	// Для таймера шага
	tonStepTimeout   : TON; // Таймер превышения времени шага
	xStepTimeout     : BOOL; // Время шага превышено
	xStepChanged     : BOOL; // Шаг изменился в текущем цикле
	xStepTimerEnable : BOOL; // Разрешение таймера шага
	xStepInitialized : BOOL; // Предыдущий шаг инициализирован
	
	// Для удержания предупреждений
    tpWarningHold : TP; // Удержание предупреждения для отображения
    xWarningPulse : BOOL; // Импульс нового предупреждения
	
	// ФБ группы осей
	fbReadStatus   : MC_GroupReadStatus; // Чтение состояния группы
	fbReadError    : MC_GroupReadError; // Чтение активной ошибки группы
	fbReadPosition : MC_GroupReadActualPosition; // Чтение текущей позиции группы
	fbGroupEnable  : MC_GroupEnable; // Включение группы
	fbGroupDisable : MC_GroupDisable; // Отключение группы
	fbGroupReset   : MC_GroupReset; // Сброс ошибок группы
	fbGroupSetOverride : MC_GroupSetOverride; // Live override активного и следующего движения группы

	
	fbMoveDirect : MC_MoveDirectAbsolute; // Прямое абсолютное перемещение
	fbMoveLinear : MC_MoveLinearAbsolute; // Линейное абсолютное перемещение
	fbFaultInjector : FB_AXIS_GROUP_FAULT_INJECTOR; // Изолированная инъекция библиотечной ошибки
	
	fbGroupHalt : MC_GroupHalt; // Плавная остановка группы
	fbGroupStop : MC_GroupStop; // Остановка группы
	
	stPosition : SMC_POS_REF; // Текущая позиция группы
	
	// Триггеры на команды
    rtEnable        : R_TRIG; // Фронт команды включения
    rtDisable       : R_TRIG; // Фронт команды отключения
	rtEnablePower   : R_TRIG; // Фронт запроса питания
    rtResetAllError : R_TRIG; // Фронт команды сброса
    rtMoveDirect    : R_TRIG; // Фронт прямого перемещения
    rtMoveLinear    : R_TRIG; // Фронт линейного перемещения
	rtStopCmd       : R_TRIG; // Фронт команды остановки
	rtHaltCmd       : R_TRIG; // Фронт плавной остановки
	
END_VAR
VAR_IN_OUT
	AxisGroup : AXIS_GROUP_REF_SM3; // Ссылка на группу осей SoftMotion
	GroupData : ST_AXIS_GROUP; // Команды, статусы и диагностика группы
END_VAR

VAR CONSTANT
	// ==================================================
    // Логические ошибки группы
    // ==================================================
	LOG_STEP_TIMEOUT             : DWORD := 1; // Превышено время шага
	LOG_INVALID_STATE            : DWORD := 2; // Неизвестный шаг автомата
	LOG_POWER_PERMIT_READY       : DWORD := 4; // Нет разрешения питания в готовности
	LOG_POWER_PERMIT_LOST_DIRECT : DWORD := 8; // Разрешение питания снято при движении
	// ==================================================
    // Ошибки блоков движения группы
    // ==================================================
	MOTION_ERR_ENABLE        : DWORD := 1; // Ошибка включения группы
	MOTION_ERR_DISABLE       : DWORD := 4; // Ошибка отключения группы
	MOTION_ERR_RESET         : DWORD := 8; // Ошибка сброса группы
	MOTION_ERR_MOVE_DIRECT   : DWORD := 16; // Ошибка прямого перемещения
	MOTION_ERR_MOVE_LINEAR   : DWORD := 32; // Ошибка линейного перемещения
	MOTION_ERR_HALT          : DWORD := 64; // Ошибка плавной остановки
	MOTION_ERR_STOP          : DWORD := 128; // Ошибка остановки
	MOTION_ERR_READ_POSITION : DWORD := 256; // Ошибка чтения позиции
	MOTION_ERR_READ_STATUS   : DWORD := 512; // Ошибка чтения статуса
	MOTION_ERR_READ_GROUP_ERROR : DWORD := 1024; // Ошибка чтения кода ошибки группы
	MOTION_ERR_GROUP_ERROR_STOP : DWORD := 2048; // Группа SoftMotion находится в ErrorStop
	MOTION_ERR_SIMULATED        : DWORD := 4096; // Тестовая ошибка MC_MoveDirectAbsolute
	MOTION_ERR_OVERRIDE         : DWORD := 8192; // Ошибка MC_GroupSetOverride; бит 1 сохранён за legacy POWER_ERROR

	WRN_NO_POWER_PERMIT       : UINT := 1; // Нет разрешения питания
	WRN_MOVE_COMMAND_CONFLICT : UINT := 2; // Одновременно заданы два типа движения
	WRN_GLOBAL_ERROR_ACTIVE   : UINT := 3; // Сброс отклонён из-за глобальной ошибки
	WRN_MOTION_ERROR_ACTIVE   : UINT := 4; // Сброс отклонён из-за активной Motion-ошибки
	WRN_RESET_VERIFY_TIMEOUT  : UINT := 5; // Не получено подтверждение сброса за допустимое время
	WRN_GROUP_ERROR_AFTER_RESET : UINT := 6; // Группа осталась в ErrorStop после сброса
	WRN_GROUP_RESET_ERROR     : UINT := 7; // MC_GroupReset завершился ошибкой
	WRN_GROUP_RESET_TIMEOUT   : UINT := 8; // Превышено время выполнения MC_GroupReset
	WRN_SIM_ERROR_NOT_ALLOWED : UINT := 9; // Тестовая ошибка запрещена текущим состоянием группы
END_VAR

// Коэффициент симуляции не изменяет динамику группы осей робота.
lrAppliedVelocityOverride := MAX(0.001, MIN(1.0, lrVelocityOverride));

// =============================================================================
// 1. Добить предупреждения и ошибки
// 2. Сделать логирование ошибок и шагов
// 3. Сделать необходимые сигналы статусов
// =============================================================================

// =============================================================================
// 1. Одноцикловые сигналы
// =============================================================================
xWarningPulse := FALSE;

GroupData.Diag.xStepChanged := FALSE;
GroupData.Error.dwLogicalErrorNew := DWORD#0;
GroupData.Error.dwMotionErrorNew := DWORD#0;


// =============================================================================
// 2. Фронты команд
// =============================================================================
rtDisable(CLK := GroupData.Command.xDisable);
rtEnablePower(CLK := GroupData.Command.xPowerEnable);
rtResetAllError(CLK := GroupData.Command.xReset);
rtMoveDirect(CLK := GroupData.Command.xMoveDirect);
rtMoveLinear(CLK := GroupData.Command.xMoveLinear);
rtHaltCmd(CLK := GroupData.Command.xHaltCmd);
rtStopCmd(CLK := GroupData.Command.xStopCmd);


// =============================================================================
// 3. Чтение состояния группы и координат
// =============================================================================
fbReadStatus(
    Enable    := TRUE,
    AxisGroup := AxisGroup
);

fbReadError(
    Enable    := TRUE,
    AxisGroup := AxisGroup
);

fbReadPosition(
    AxisGroup   := AxisGroup,
    Enable      := TRUE,
    CoordSystem := SMC_COORD_SYSTEM.MCS
);

IF fbReadPosition.Valid THEN
	stPosition := fbReadPosition.Position;
    GroupData.Status.ActualX := fbReadPosition.Position.c.X;
    GroupData.Status.ActualY := fbReadPosition.Position.c.Y;
    GroupData.Status.ActualZ := fbReadPosition.Position.c.Z;
END_IF;
GroupData.Status.xPositionValid := fbReadPosition.Valid AND NOT fbReadPosition.Error;


// =============================================================================
// 4. Текущий статус ошибок
// =============================================================================
GroupData.Status.xGroupError :=
    fbReadStatus.Error
    OR fbReadStatus.GroupErrorStop
    OR (GroupData.Error.dwMotionErrorLatched <> DWORD#0);

GroupData.Status.xLogicalError :=
    GroupData.Error.dwLogicalErrorLatched <> DWORD#0;

GroupData.Status.xLocalError :=
    GroupData.Status.xGroupError
    OR GroupData.Status.xLogicalError;

// Тестовый Motion-FB запускается только в неподвижной готовой группе.
xFaultAllowed := fbReadStatus.Valid
	AND fbReadStatus.GroupStandby
	AND (GroupData.Diag.iStep = E_AXIS_GROUP_STATE.READY)
	AND NOT GroupData.Status.xLocalError
	AND NOT GroupData.Command.xGlobalError
	AND NOT GroupData.Command.xMoveDirect
	AND NOT GroupData.Command.xMoveLinear;

fbFaultInjector(
	Request := FaultRequest,
	xOwnerAllowed := xFaultAllowed,
	xReset := GroupData.Command.xReset,
	Position := stPosition,
	AxisGroup := AxisGroup
);
FaultStatus := fbFaultInjector.Status;

IF fbFaultInjector.Status.xRejected THEN
	GroupData.Diag.sWarningText := 'Simulated SM3 error is not allowed';
	GroupData.Diag.stWarning.uiCode := WRN_SIM_ERROR_NOT_ALLOWED;
	GroupData.Diag.stWarning.udiSequence := GroupData.Diag.stWarning.udiSequence + UDINT#1;
	IF GroupData.Diag.stWarning.udiSequence = UDINT#0 THEN
		GroupData.Diag.stWarning.udiSequence := UDINT#1;
	END_IF;
	xWarningPulse := TRUE;
END_IF;


// =============================================================================
// 5. Команды Motion FB по умолчанию
// =============================================================================
xEnable := FALSE;
xDisable := FALSE;
xResetMC := FALSE;
xMoveDirect := FALSE;
xMoveLinear := FALSE;
xStopCmd := FALSE;
xHaltCmd := FALSE;


// =============================================================================
// 6. Машина состояний
// =============================================================================
CASE GroupData.Diag.iStep OF

    // -------------------------------------------------------------------------
    E_AXIS_GROUP_STATE.DISABLED:
    // -------------------------------------------------------------------------
        GroupData.Diag.sStepName := 'DISABLED';
        GroupData.Diag.tStepPreset := T#0S;
        GroupData.Diag.iPowerMode := E_AXIS_GROUP_POWER_MODE.OFF;

        IF GroupData.Command.xGlobalError
           OR GroupData.Status.xLocalError THEN

            GroupData.Diag.iStep := E_AXIS_GROUP_STATE.ERROR;

        ELSIF rtEnablePower.Q AND NOT GroupData.Command.xPowerPermit THEN
            GroupData.Diag.sWarningText := 'Power permit is not active';
            GroupData.Diag.stWarning.uiCode := WRN_NO_POWER_PERMIT;
            GroupData.Diag.stWarning.udiSequence := GroupData.Diag.stWarning.udiSequence + UDINT#1;
            IF GroupData.Diag.stWarning.udiSequence = UDINT#0 THEN
                GroupData.Diag.stWarning.udiSequence := UDINT#1;
            END_IF;
            xWarningPulse := TRUE;

		ELSIF fbReadStatus.Valid AND fbReadStatus.GroupStandby THEN
			// MC_GroupReset всегда возвращает группу в GroupStandby. Если питание
			// запрошено, используем это состояние без повторного MC_GroupEnable;
			// иначе сначала синхронизируем группу с программным шагом DISABLED.
			IF rtEnablePower.Q THEN
				GroupData.Diag.iStep := E_AXIS_GROUP_STATE.ENABLING_POWER;
			ELSE
				GroupData.Diag.iStep := E_AXIS_GROUP_STATE.DISABLING_GROUP;
			END_IF;

        ELSIF rtEnablePower.Q THEN
            GroupData.Diag.iStep := E_AXIS_GROUP_STATE.ENABLING_POWER;
        END_IF;


    // -------------------------------------------------------------------------
    E_AXIS_GROUP_STATE.ENABLING_POWER:
    // -------------------------------------------------------------------------
        GroupData.Diag.sStepName := 'ENABLING_POWER';
        GroupData.Diag.tStepPreset := GroupData.Timeouts.tPowerTimeout;
        GroupData.Diag.iPowerMode := E_AXIS_GROUP_POWER_MODE.ON;

        IF fbReadStatus.GroupErrorStop THEN

            GroupData.Diag.iStep := E_AXIS_GROUP_STATE.ERROR;

        ELSIF NOT GroupData.Command.xPowerPermit
           OR GroupData.Command.xGlobalError THEN

            GroupData.Diag.iStep := E_AXIS_GROUP_STATE.DISABLING_POWER;

        ELSIF xStepTimeout THEN
            GroupData.Error.dwLogicalErrorNew :=
                GroupData.Error.dwLogicalErrorNew
                OR LOG_STEP_TIMEOUT;

            GroupData.Diag.iStep := E_AXIS_GROUP_STATE.DISABLING_POWER;

		ELSIF xAxesPowered AND fbReadStatus.Valid THEN
			IF fbReadStatus.GroupStandby THEN
				GroupData.Diag.iStep := E_AXIS_GROUP_STATE.READY;
			ELSIF fbReadStatus.GroupDisabled THEN
				GroupData.Diag.iStep := E_AXIS_GROUP_STATE.ENABLING_GROUP;
			END_IF;
		END_IF;


    // -------------------------------------------------------------------------
    E_AXIS_GROUP_STATE.ENABLING_GROUP:
    // -------------------------------------------------------------------------
        GroupData.Diag.sStepName := 'ENABLING_GROUP';
        GroupData.Diag.tStepPreset := GroupData.Timeouts.tGroupTimeout;
        GroupData.Diag.iPowerMode := E_AXIS_GROUP_POWER_MODE.ON;

		// MC_GroupEnable допустим только из GroupDisabled. Execute формируется
		// исключительно на этом шаге: после перехода в GroupStandby он снимается,
		// чтобы новый фронт не вызвал MC_GroupEnable повторно после MC_GroupReset.
		xEnable := fbReadStatus.Valid AND fbReadStatus.GroupDisabled;

		IF fbReadStatus.GroupErrorStop THEN

            GroupData.Diag.iStep := E_AXIS_GROUP_STATE.ERROR;

		ELSIF fbReadStatus.Valid AND fbReadStatus.GroupStandby THEN

			GroupData.Diag.iStep := E_AXIS_GROUP_STATE.READY;

		ELSIF xEnable AND fbGroupEnable.Error THEN

			GroupData.Diag.iStep := E_AXIS_GROUP_STATE.ERROR;

        ELSIF NOT GroupData.Command.xPowerPermit
           OR GroupData.Command.xGlobalError THEN

            GroupData.Diag.iStep := E_AXIS_GROUP_STATE.DISABLING_GROUP;

        ELSIF xStepTimeout THEN
            GroupData.Error.dwLogicalErrorNew :=
                GroupData.Error.dwLogicalErrorNew
                OR LOG_STEP_TIMEOUT;

            GroupData.Diag.iStep := E_AXIS_GROUP_STATE.DISABLING_GROUP;

		END_IF;


    // -------------------------------------------------------------------------
    E_AXIS_GROUP_STATE.READY:
    // -------------------------------------------------------------------------
        GroupData.Diag.sStepName := 'READY';
        GroupData.Diag.tStepPreset := T#0S;
        GroupData.Diag.iPowerMode := E_AXIS_GROUP_POWER_MODE.ON;

		IF fbReadStatus.GroupErrorStop THEN
            GroupData.Diag.iStep := E_AXIS_GROUP_STATE.ERROR;

        ELSIF NOT GroupData.Command.xPowerPermit
           OR GroupData.Command.xGlobalError
           OR GroupData.Status.xLocalError
           OR rtDisable.Q THEN

            GroupData.Diag.iStep := E_AXIS_GROUP_STATE.DISABLING_GROUP;

        ELSIF rtMoveDirect.Q AND rtMoveLinear.Q THEN
            GroupData.Diag.sWarningText :=
                'MoveDirect and MoveLinear requested together';

            GroupData.Diag.stWarning.uiCode := WRN_MOVE_COMMAND_CONFLICT;
            GroupData.Diag.stWarning.udiSequence := GroupData.Diag.stWarning.udiSequence + UDINT#1;
            IF GroupData.Diag.stWarning.udiSequence = UDINT#0 THEN
                GroupData.Diag.stWarning.udiSequence := UDINT#1;
            END_IF;

            xWarningPulse := TRUE;

        ELSIF rtMoveDirect.Q THEN
            GroupData.Diag.iStep := E_AXIS_GROUP_STATE.MOVING_DIRECT;

        ELSIF rtMoveLinear.Q THEN
            GroupData.Diag.iStep := E_AXIS_GROUP_STATE.MOVING_LINEAR;
        END_IF;


    // -------------------------------------------------------------------------
    E_AXIS_GROUP_STATE.MOVING_DIRECT:
    // -------------------------------------------------------------------------
        GroupData.Diag.sStepName := 'MOVING_DIRECT';
        GroupData.Diag.tStepPreset := GroupData.Timeouts.tMoveTimeout;
        GroupData.Diag.iPowerMode := E_AXIS_GROUP_POWER_MODE.ON;

		xMoveDirect := TRUE;

        IF fbReadStatus.GroupErrorStop THEN
            GroupData.Diag.iStep := E_AXIS_GROUP_STATE.ERROR;

        ELSIF fbMoveDirect.Error THEN
            IF fbReadStatus.GroupMoving THEN
                GroupData.Diag.iStep := E_AXIS_GROUP_STATE.EMG_STOP;
            ELSE
                GroupData.Diag.iStep := E_AXIS_GROUP_STATE.ERROR;
            END_IF;

        ELSIF xStepTimeout THEN
            GroupData.Error.dwLogicalErrorNew :=
                GroupData.Error.dwLogicalErrorNew
                OR LOG_STEP_TIMEOUT;

            GroupData.Diag.iStep := E_AXIS_GROUP_STATE.EMG_STOP;

        ELSIF NOT GroupData.Command.xPowerPermit
           OR GroupData.Command.xGlobalError
           OR GroupData.Status.xLocalError
           OR rtStopCmd.Q THEN

            GroupData.Diag.iStep := E_AXIS_GROUP_STATE.EMG_STOP;

        ELSIF rtHaltCmd.Q THEN
            GroupData.Diag.iStep := E_AXIS_GROUP_STATE.HALT_STOP;

        ELSIF fbMoveDirect.Done
           AND fbReadStatus.GroupStandby THEN

            GroupData.Diag.iStep := E_AXIS_GROUP_STATE.READY;
        END_IF;

    // -------------------------------------------------------------------------
    E_AXIS_GROUP_STATE.HALT_STOP:
    // -------------------------------------------------------------------------
        GroupData.Diag.sStepName := 'HALT_STOP';
        GroupData.Diag.tStepPreset := GroupData.Timeouts.tHaltTimeout;
        GroupData.Diag.iPowerMode := E_AXIS_GROUP_POWER_MODE.ON;

		xHaltCmd := TRUE;

        IF fbReadStatus.GroupErrorStop THEN
            GroupData.Diag.iStep := E_AXIS_GROUP_STATE.ERROR;

        ELSIF fbGroupHalt.Error
           OR xStepTimeout
           OR NOT GroupData.Command.xPowerPermit
           OR GroupData.Command.xGlobalError
           OR GroupData.Status.xLocalError
           OR rtStopCmd.Q THEN

            IF xStepTimeout THEN
                GroupData.Error.dwLogicalErrorNew :=
                    GroupData.Error.dwLogicalErrorNew
                    OR LOG_STEP_TIMEOUT;
            END_IF;

            GroupData.Diag.iStep := E_AXIS_GROUP_STATE.EMG_STOP;

        ELSIF fbGroupHalt.Done
           AND fbReadStatus.GroupStandby THEN

            GroupData.Diag.iStep := E_AXIS_GROUP_STATE.READY;
        END_IF;


    // -------------------------------------------------------------------------
    E_AXIS_GROUP_STATE.EMG_STOP:
    // -------------------------------------------------------------------------
        GroupData.Diag.sStepName := 'STOPPING';
        GroupData.Diag.tStepPreset := GroupData.Timeouts.tStopTimeout;
        GroupData.Diag.iPowerMode := E_AXIS_GROUP_POWER_MODE.ON;

		xStopCmd := TRUE;

        IF fbReadStatus.GroupErrorStop
           OR fbGroupStop.Error THEN

            GroupData.Diag.iStep := E_AXIS_GROUP_STATE.ERROR;

        ELSIF xStepTimeout THEN
            GroupData.Error.dwLogicalErrorNew :=
                GroupData.Error.dwLogicalErrorNew
                OR LOG_STEP_TIMEOUT;

            GroupData.Diag.iStep := E_AXIS_GROUP_STATE.ERROR;

        ELSIF fbGroupStop.Done THEN
            GroupData.Diag.iStep := E_AXIS_GROUP_STATE.WAIT_STOP;
        END_IF;


    // -------------------------------------------------------------------------
    E_AXIS_GROUP_STATE.WAIT_STOP:
    // -------------------------------------------------------------------------
        GroupData.Diag.sStepName := 'WAIT_STOP';
        GroupData.Diag.tStepPreset := GroupData.Timeouts.tStopTimeout;
        GroupData.Diag.iPowerMode := E_AXIS_GROUP_POWER_MODE.ON;

		IF fbReadStatus.GroupErrorStop THEN
            GroupData.Diag.iStep := E_AXIS_GROUP_STATE.ERROR;

        ELSIF xStepTimeout THEN
            GroupData.Error.dwLogicalErrorNew :=
                GroupData.Error.dwLogicalErrorNew
                OR LOG_STEP_TIMEOUT;

            GroupData.Diag.iStep := E_AXIS_GROUP_STATE.ERROR;

		ELSIF fbReadStatus.GroupStandby THEN
			// Операторский Stop завершает только движение и сохраняет GroupStandby.
			// Отключение группы выполняется лишь по отдельному запросу питания/ошибке.
			IF GroupData.Command.xPowerPermit
			AND NOT GroupData.Command.xDisable
			AND NOT GroupData.Command.xGlobalError
			AND NOT GroupData.Status.xLocalError THEN
				GroupData.Diag.iStep := E_AXIS_GROUP_STATE.READY;
			ELSE
				GroupData.Diag.iStep := E_AXIS_GROUP_STATE.DISABLING_GROUP;
			END_IF;
		END_IF;


    // -------------------------------------------------------------------------
    E_AXIS_GROUP_STATE.DISABLING_GROUP:
    // -------------------------------------------------------------------------
        GroupData.Diag.sStepName := 'DISABLING_GROUP';
        GroupData.Diag.tStepPreset := GroupData.Timeouts.tGroupTimeout;
        GroupData.Diag.iPowerMode := E_AXIS_GROUP_POWER_MODE.ON;

		// MC_GroupDisable допустим только из GroupStandby.
		xDisable := fbReadStatus.Valid AND fbReadStatus.GroupStandby;

		IF fbReadStatus.GroupErrorStop THEN

            GroupData.Diag.iStep := E_AXIS_GROUP_STATE.ERROR;

		ELSIF fbReadStatus.Valid AND fbReadStatus.GroupDisabled THEN

			GroupData.Diag.iStep := E_AXIS_GROUP_STATE.DISABLING_POWER;

		ELSIF xDisable AND fbGroupDisable.Error THEN

			GroupData.Diag.iStep := E_AXIS_GROUP_STATE.ERROR;

        ELSIF xStepTimeout THEN
            GroupData.Error.dwLogicalErrorNew :=
                GroupData.Error.dwLogicalErrorNew
                OR LOG_STEP_TIMEOUT;

            GroupData.Diag.iStep := E_AXIS_GROUP_STATE.ERROR;

		ELSIF xDisable AND fbGroupDisable.Done
           AND fbReadStatus.GroupDisabled THEN

            GroupData.Diag.iStep := E_AXIS_GROUP_STATE.DISABLING_POWER;
        END_IF;


    // -------------------------------------------------------------------------
    E_AXIS_GROUP_STATE.DISABLING_POWER:
    // -------------------------------------------------------------------------
        GroupData.Diag.sStepName := 'DISABLING_POWER';
        GroupData.Diag.tStepPreset := GroupData.Timeouts.tPowerTimeout;
        GroupData.Diag.iPowerMode :=
            E_AXIS_GROUP_POWER_MODE.OFF_REQUEST;

        IF xStepTimeout THEN
            GroupData.Error.dwLogicalErrorNew :=
                GroupData.Error.dwLogicalErrorNew
                OR LOG_STEP_TIMEOUT;

            GroupData.Diag.iStep := E_AXIS_GROUP_STATE.ERROR;

        ELSIF NOT xAxesPowered THEN

            IF GroupData.Command.xGlobalError
               OR GroupData.Status.xLocalError
			   OR NOT GroupData.Command.xPowerPermit THEN

                GroupData.Diag.iStep := E_AXIS_GROUP_STATE.ERROR;
            ELSE
                GroupData.Diag.iStep := E_AXIS_GROUP_STATE.DISABLED;
            END_IF;
        END_IF;


    // -------------------------------------------------------------------------
    E_AXIS_GROUP_STATE.ERROR:
    // -------------------------------------------------------------------------
        GroupData.Diag.sStepName := 'ERROR';
        GroupData.Diag.tStepPreset := T#0S;

        GroupData.Diag.iPowerMode := E_AXIS_GROUP_POWER_MODE.OFF_REQUEST;

		IF rtResetAllError.Q AND xResetPermit THEN

            IF GroupData.Command.xGlobalError THEN
                GroupData.Diag.sWarningText :=
                    'Global error is still active';

                GroupData.Diag.stWarning.uiCode := WRN_GLOBAL_ERROR_ACTIVE;
                GroupData.Diag.stWarning.udiSequence := GroupData.Diag.stWarning.udiSequence + UDINT#1;
                IF GroupData.Diag.stWarning.udiSequence = UDINT#0 THEN
                    GroupData.Diag.stWarning.udiSequence := UDINT#1;
                END_IF;

                xWarningPulse := TRUE;

            ELSIF fbReadStatus.GroupErrorStop THEN
                    GroupData.Diag.iStep :=
                        E_AXIS_GROUP_STATE.RESETTING;

            ELSIF GroupData.Error.dwMotionErrorActive
                  <> DWORD#0 THEN

                GroupData.Diag.sWarningText :=
                    'Motion FB error is still active';

                GroupData.Diag.stWarning.uiCode := WRN_MOTION_ERROR_ACTIVE;
                GroupData.Diag.stWarning.udiSequence := GroupData.Diag.stWarning.udiSequence + UDINT#1;
                IF GroupData.Diag.stWarning.udiSequence = UDINT#0 THEN
                    GroupData.Diag.stWarning.udiSequence := UDINT#1;
                END_IF;

                xWarningPulse := TRUE;

            ELSE
                // Ошибка устранена — очищаем защёлки.
                GroupData.Error.dwLogicalErrorLatched := DWORD#0;
                GroupData.Error.dwMotionErrorLatched := DWORD#0;
                GroupData.Error.dwMotionErrorPrevious := DWORD#0;

				IF fbReadStatus.GroupStandby AND NOT xAxesPowered THEN
					GroupData.Diag.iStep :=
						E_AXIS_GROUP_STATE.DISABLING_GROUP;

				ELSIF fbReadStatus.GroupDisabled AND NOT xAxesPowered THEN
					GroupData.Diag.iStep :=
						E_AXIS_GROUP_STATE.DISABLED;

				ELSIF fbReadStatus.GroupDisabled THEN
					GroupData.Diag.iStep :=
						E_AXIS_GROUP_STATE.ENABLING_GROUP;

                ELSIF fbReadStatus.GroupStandby THEN
                    GroupData.Diag.iStep :=
                        E_AXIS_GROUP_STATE.READY;

                ELSE
                    GroupData.Diag.iStep :=
                        E_AXIS_GROUP_STATE.DISABLING_POWER;
                END_IF;
            END_IF;
        END_IF;


    // -------------------------------------------------------------------------
    E_AXIS_GROUP_STATE.RESETTING:
    // -------------------------------------------------------------------------
        GroupData.Diag.sStepName := 'RESETTING';
        GroupData.Diag.tStepPreset := GroupData.Timeouts.tGroupTimeout;
        GroupData.Diag.iPowerMode := E_AXIS_GROUP_POWER_MODE.ON;

		// Ошибка оси могла исчезнуть между принятием общей команды и этим циклом.
		// В таком случае MC_GroupReset не вызывается, иначе он вернёт 78
		// (no error to be resetted); остаётся только очистить внутренние защёлки.
		IF fbReadStatus.Valid AND NOT fbReadStatus.GroupErrorStop THEN
			xResetMC := FALSE;
			GroupData.Diag.iStep := E_AXIS_GROUP_STATE.RESET_VERIFY;

		ELSE
			xResetMC := TRUE;
		END_IF;

		IF GroupData.Command.xGlobalError THEN
            GroupData.Diag.sWarningText :=
                'Global error became active during group reset';

            GroupData.Diag.stWarning.uiCode := WRN_GLOBAL_ERROR_ACTIVE;
            GroupData.Diag.stWarning.udiSequence := GroupData.Diag.stWarning.udiSequence + UDINT#1;
            IF GroupData.Diag.stWarning.udiSequence = UDINT#0 THEN
                GroupData.Diag.stWarning.udiSequence := UDINT#1;
            END_IF;

            xWarningPulse := TRUE;
            GroupData.Diag.iStep := E_AXIS_GROUP_STATE.ERROR;

		ELSIF xResetMC AND fbGroupReset.Error THEN
            GroupData.Diag.sWarningText :=
                'MC_GroupReset finished with error';

            GroupData.Diag.stWarning.uiCode := WRN_GROUP_RESET_ERROR;
            GroupData.Diag.stWarning.udiSequence := GroupData.Diag.stWarning.udiSequence + UDINT#1;
            IF GroupData.Diag.stWarning.udiSequence = UDINT#0 THEN
                GroupData.Diag.stWarning.udiSequence := UDINT#1;
            END_IF;

            xWarningPulse := TRUE;
            GroupData.Diag.iStep := E_AXIS_GROUP_STATE.ERROR;

		ELSIF xResetMC AND xStepTimeout THEN
            GroupData.Diag.sWarningText :=
                'MC_GroupReset timeout';

            GroupData.Diag.stWarning.uiCode := WRN_GROUP_RESET_TIMEOUT;
            GroupData.Diag.stWarning.udiSequence := GroupData.Diag.stWarning.udiSequence + UDINT#1;
            IF GroupData.Diag.stWarning.udiSequence = UDINT#0 THEN
                GroupData.Diag.stWarning.udiSequence := UDINT#1;
            END_IF;

            xWarningPulse := TRUE;
            GroupData.Error.dwLogicalErrorNew :=
                GroupData.Error.dwLogicalErrorNew
                OR LOG_STEP_TIMEOUT;

            GroupData.Diag.iStep := E_AXIS_GROUP_STATE.ERROR;

		ELSIF xResetMC AND fbGroupReset.Done THEN
            // Статус группы был прочитан до вызова MC_GroupReset.
            // Проверяем результат сброса только со следующего цикла.
            GroupData.Diag.iStep := E_AXIS_GROUP_STATE.RESET_VERIFY;
        END_IF;


    // -------------------------------------------------------------------------
    E_AXIS_GROUP_STATE.RESET_VERIFY:
    // -------------------------------------------------------------------------
        GroupData.Diag.sStepName := 'RESET_VERIFY';
        GroupData.Diag.tStepPreset := GroupData.Timeouts.tGroupTimeout;
        GroupData.Diag.iPowerMode := E_AXIS_GROUP_POWER_MODE.ON;

        IF GroupData.Command.xGlobalError THEN
            GroupData.Diag.sWarningText :=
                'Global error became active during reset verification';

            GroupData.Diag.stWarning.uiCode := WRN_GLOBAL_ERROR_ACTIVE;
            GroupData.Diag.stWarning.udiSequence := GroupData.Diag.stWarning.udiSequence + UDINT#1;
            IF GroupData.Diag.stWarning.udiSequence = UDINT#0 THEN
                GroupData.Diag.stWarning.udiSequence := UDINT#1;
            END_IF;

            xWarningPulse := TRUE;
            GroupData.Diag.iStep := E_AXIS_GROUP_STATE.ERROR;

        ELSIF xStepTimeout THEN
            GroupData.Diag.sWarningText :=
                'Reset verification timeout';

            GroupData.Diag.stWarning.uiCode := WRN_RESET_VERIFY_TIMEOUT;
            GroupData.Diag.stWarning.udiSequence := GroupData.Diag.stWarning.udiSequence + UDINT#1;
            IF GroupData.Diag.stWarning.udiSequence = UDINT#0 THEN
                GroupData.Diag.stWarning.udiSequence := UDINT#1;
            END_IF;

            xWarningPulse := TRUE;
            GroupData.Error.dwLogicalErrorNew :=
                GroupData.Error.dwLogicalErrorNew
                OR LOG_STEP_TIMEOUT;

            GroupData.Diag.iStep := E_AXIS_GROUP_STATE.ERROR;

        ELSIF fbReadStatus.Valid
           AND fbReadStatus.GroupErrorStop
           AND fbReadError.Valid
           AND (TO_UDINT(fbReadError.GroupErrorID) <> UDINT#0) THEN

            // Причина ошибки осталась активной после завершения сброса.
            GroupData.Diag.sWarningText :=
                'Axis group error remains active after reset';

            GroupData.Diag.stWarning.uiCode := WRN_GROUP_ERROR_AFTER_RESET;
            GroupData.Diag.stWarning.udiSequence := GroupData.Diag.stWarning.udiSequence + UDINT#1;
            IF GroupData.Diag.stWarning.udiSequence = UDINT#0 THEN
                GroupData.Diag.stWarning.udiSequence := UDINT#1;
            END_IF;

            xWarningPulse := TRUE;
            GroupData.Diag.iStep := E_AXIS_GROUP_STATE.ERROR;

        ELSIF fbReadStatus.Valid
           AND NOT fbReadStatus.GroupErrorStop THEN

            GroupData.Error.dwLogicalErrorLatched := DWORD#0;
            GroupData.Error.dwMotionErrorLatched := DWORD#0;
            GroupData.Error.dwMotionErrorPrevious := DWORD#0;

			IF fbReadStatus.GroupStandby AND NOT xAxesPowered THEN
				GroupData.Diag.iStep := E_AXIS_GROUP_STATE.DISABLING_GROUP;

			ELSIF fbReadStatus.GroupDisabled AND NOT xAxesPowered THEN
				GroupData.Diag.iStep := E_AXIS_GROUP_STATE.DISABLED;

			ELSIF fbReadStatus.GroupDisabled THEN
				GroupData.Diag.iStep := E_AXIS_GROUP_STATE.ENABLING_GROUP;

            ELSIF fbReadStatus.GroupStandby THEN
                GroupData.Diag.iStep := E_AXIS_GROUP_STATE.READY;

            ELSE
                GroupData.Diag.iStep := E_AXIS_GROUP_STATE.DISABLING_POWER;
            END_IF;
        END_IF;


    // -------------------------------------------------------------------------
    ELSE
    // -------------------------------------------------------------------------
        GroupData.Error.dwLogicalErrorNew :=
            GroupData.Error.dwLogicalErrorNew
            OR LOG_INVALID_STATE;

        GroupData.Diag.iStep := E_AXIS_GROUP_STATE.ERROR;

END_CASE;


// =============================================================================
// 7. Целевая позиция
// =============================================================================
GroupData.MotionParam.stTargetPos.c.X := GroupData.MotionParam.lrX;
GroupData.MotionParam.stTargetPos.c.Y := GroupData.MotionParam.lrY;
GroupData.MotionParam.stTargetPos.c.Z := GroupData.MotionParam.lrZ;


// =============================================================================
// 8. Вызовы Motion FB
// =============================================================================
fbGroupEnable(
    AxisGroup := AxisGroup,
    Execute   := xEnable
);

fbGroupDisable(
    AxisGroup := AxisGroup,
    Execute   := xDisable
);

fbGroupReset(
    AxisGroup := AxisGroup,
    Execute   := xResetMC
);

// MC_GroupSetOverride меняет скорость уже активного движения. Вызов обязан
// находиться перед Motion FB. Во время MC_GroupStop блок запрещён документацией:
// последняя записанная величина сохраняется, а Stop выполняется со своей динамикой.
xVelocityOverrideEnable := fbReadStatus.Valid
	AND NOT fbReadStatus.GroupErrorStop
	AND NOT xStopCmd
	AND ((GroupData.Diag.iStep = E_AXIS_GROUP_STATE.READY)
		OR (GroupData.Diag.iStep = E_AXIS_GROUP_STATE.MOVING_DIRECT)
		OR (GroupData.Diag.iStep = E_AXIS_GROUP_STATE.MOVING_LINEAR));
fbGroupSetOverride(
	AxisGroup      := AxisGroup,
	Enable         := xVelocityOverrideEnable,
	VelFactor      := lrAppliedVelocityOverride,
	AccFactor      := 1.0,
	JerkFactor     := 1.0,
	TorqueFactor   := 1.0,
	PathVelFactor  := lrAppliedVelocityOverride,
	PathAccFactor  := 1.0,
	PathJerkFactor := 1.0
);

fbMoveDirect(
    AxisGroup   := AxisGroup,
    Execute     := xMoveDirect,
    Position    := GroupData.MotionParam.stTargetPos,
    CoordSystem := SMC_COORD_SYSTEM.MCS,
    BufferMode  := MC_BUFFER_MODE.Aborting,
	// Коэффициент точки задаёт профиль команды, общий процент накладывается
	// отдельно через MC_GroupSetOverride и потому здесь повторно не умножается.
	VelFactor   := MAX(0.001, MIN(1.0, GroupData.MotionParam.VelFactor)),
    AccFactor   := GroupData.MotionParam.AccFactor,
    JerkFactor  := GroupData.MotionParam.JerkFactor
);

fbMoveLinear(
    AxisGroup := AxisGroup,
    Execute   := xMoveLinear
);

fbGroupHalt(
	AxisGroup    := AxisGroup,
	Execute      := xHaltCmd,
	Deceleration := GroupData.MotionParam.HaltDeceleration,
	Jerk         := GroupData.MotionParam.HaltJerk
);

fbGroupStop(
	AxisGroup    := AxisGroup,
	Execute      := xStopCmd,
	Deceleration := GroupData.MotionParam.HaltDeceleration * 2,
	Jerk         := GroupData.MotionParam.HaltJerk * 2
);


// =============================================================================
// 9. Маска Motion-ошибок
// =============================================================================
GroupData.Error.dwMotionErrorActive := DWORD#0;

IF fbGroupEnable.Error THEN
    GroupData.Error.dwMotionErrorActive :=
        GroupData.Error.dwMotionErrorActive
        OR MOTION_ERR_ENABLE;
END_IF;

IF fbGroupDisable.Error THEN
    GroupData.Error.dwMotionErrorActive :=
        GroupData.Error.dwMotionErrorActive
        OR MOTION_ERR_DISABLE;
END_IF;

IF fbGroupReset.Error THEN
    GroupData.Error.dwMotionErrorActive :=
        GroupData.Error.dwMotionErrorActive
        OR MOTION_ERR_RESET;
END_IF;

IF fbMoveDirect.Error THEN
    GroupData.Error.dwMotionErrorActive :=
        GroupData.Error.dwMotionErrorActive
        OR MOTION_ERR_MOVE_DIRECT;
END_IF;

IF fbMoveLinear.Error THEN
    GroupData.Error.dwMotionErrorActive :=
        GroupData.Error.dwMotionErrorActive
        OR MOTION_ERR_MOVE_LINEAR;
END_IF;

IF fbGroupHalt.Error THEN
    GroupData.Error.dwMotionErrorActive :=
        GroupData.Error.dwMotionErrorActive
        OR MOTION_ERR_HALT;
END_IF;

IF fbGroupStop.Error THEN
    GroupData.Error.dwMotionErrorActive :=
        GroupData.Error.dwMotionErrorActive
        OR MOTION_ERR_STOP;
END_IF;

IF fbReadPosition.Error THEN
    GroupData.Error.dwMotionErrorActive :=
        GroupData.Error.dwMotionErrorActive
        OR MOTION_ERR_READ_POSITION;
END_IF;

IF fbReadStatus.Error THEN
    GroupData.Error.dwMotionErrorActive :=
        GroupData.Error.dwMotionErrorActive
        OR MOTION_ERR_READ_STATUS;
END_IF;

IF fbReadError.Error THEN
    GroupData.Error.dwMotionErrorActive :=
        GroupData.Error.dwMotionErrorActive
        OR MOTION_ERR_READ_GROUP_ERROR;
END_IF;

IF fbReadStatus.GroupErrorStop THEN
    GroupData.Error.dwMotionErrorActive :=
        GroupData.Error.dwMotionErrorActive
        OR MOTION_ERR_GROUP_ERROR_STOP;
END_IF;

IF fbFaultInjector.xError THEN
	GroupData.Error.dwMotionErrorActive :=
		GroupData.Error.dwMotionErrorActive
		OR MOTION_ERR_SIMULATED;
END_IF;

IF fbGroupSetOverride.Error THEN
	GroupData.Error.dwMotionErrorActive :=
		GroupData.Error.dwMotionErrorActive
		OR MOTION_ERR_OVERRIDE;
END_IF;

// Только ошибки, которых не было в предыдущем цикле.
GroupData.Error.dwMotionErrorNew :=
    GroupData.Error.dwMotionErrorActive
    AND NOT GroupData.Error.dwMotionErrorPrevious;


// Защёлкиваем новые логические и Motion-ошибки.
GroupData.Error.dwLogicalErrorLatched :=
    GroupData.Error.dwLogicalErrorLatched
    OR GroupData.Error.dwLogicalErrorNew;

GroupData.Error.dwMotionErrorLatched :=
    GroupData.Error.dwMotionErrorLatched
    OR GroupData.Error.dwMotionErrorNew;


// Сохраняем Motion-маску для следующего цикла.
GroupData.Error.dwMotionErrorPrevious :=
    GroupData.Error.dwMotionErrorActive;

GroupData.Error.dwAlarmActive :=
    GroupData.Error.dwMotionErrorLatched
    OR SHL(GroupData.Error.dwLogicalErrorLatched, 16);


// =============================================================================
// 11. Изменение шага и таймер
// =============================================================================
IF NOT xStepInitialized THEN
    iPrevStep := GroupData.Diag.iStep;
    xStepInitialized := TRUE;
END_IF;

xStepChanged :=
    GroupData.Diag.iStep <> iPrevStep;

GroupData.Diag.xStepChanged := xStepChanged;

IF xStepChanged THEN
    GroupData.Diag.iOldStep := iPrevStep;
    GroupData.Diag.iNewStep := GroupData.Diag.iStep;
    iPrevStep := GroupData.Diag.iStep;
END_IF;


// При переходе в новый шаг таймер один цикл выключен.
// Со следующего цикла начинается отсчёт нового шага.
tonStepTimeout(
    IN :=
        NOT xStepChanged
        AND (GroupData.Diag.tStepPreset > T#0S)
        AND (GroupData.Diag.iStep <> E_AXIS_GROUP_STATE.ERROR),

    PT := GroupData.Diag.tStepPreset
);

xStepTimeout := tonStepTimeout.Q;
GroupData.Diag.xStepTimeout := xStepTimeout;


// =============================================================================
// 12. Финальные статусы
// =============================================================================
GroupData.Status.xGroupError :=
    fbReadStatus.Error
    OR fbReadStatus.GroupErrorStop
    OR (GroupData.Error.dwMotionErrorLatched <> DWORD#0);

GroupData.Status.xLogicalError :=
    GroupData.Error.dwLogicalErrorLatched <> DWORD#0;

GroupData.Status.xLocalError :=
    GroupData.Status.xGroupError
    OR GroupData.Status.xLogicalError;

GroupData.Status.xSimErrorAllowed := FaultStatus.xAllowed;
	
GroupData.Status.xMoveDirectDone := fbMoveDirect.Done;

// Код ошибки самой группы не совпадает с ErrorID диагностических Motion FB.
IF fbReadError.Valid
   AND (TO_UDINT(fbReadError.GroupErrorID) <> UDINT#0) THEN
    GroupData.Diag.udiActualErrorID := TO_UDINT(fbReadError.GroupErrorID);
    GroupData.Diag.sErrorText := 'Axis group error';
ELSIF (GroupData.Error.dwMotionErrorLatched AND MOTION_ERR_SIMULATED) <> DWORD#0 THEN
	GroupData.Diag.udiActualErrorID := fbFaultInjector.udiErrorID;
	GroupData.Diag.sErrorText := 'Simulated MC_MoveDirectAbsolute error';
ELSIF fbGroupSetOverride.Error THEN
	GroupData.Diag.udiActualErrorID := TO_UDINT(fbGroupSetOverride.ErrorID);
	GroupData.Diag.sErrorText := 'MC_GroupSetOverride error';
ELSIF fbGroupEnable.Error THEN
	GroupData.Diag.udiActualErrorID := TO_UDINT(fbGroupEnable.ErrorID);
	GroupData.Diag.sErrorText := 'MC_GroupEnable error';
ELSIF fbGroupDisable.Error THEN
	GroupData.Diag.udiActualErrorID := TO_UDINT(fbGroupDisable.ErrorID);
	GroupData.Diag.sErrorText := 'MC_GroupDisable error';
ELSIF fbGroupReset.Error THEN
    GroupData.Diag.udiActualErrorID := TO_UDINT(fbGroupReset.ErrorID);
    GroupData.Diag.sErrorText := 'MC_GroupReset error';
ELSIF fbMoveDirect.Error THEN
	GroupData.Diag.udiActualErrorID := TO_UDINT(fbMoveDirect.ErrorID);
	GroupData.Diag.sErrorText := 'MC_MoveDirectAbsolute error';
ELSIF fbMoveLinear.Error THEN
	GroupData.Diag.udiActualErrorID := TO_UDINT(fbMoveLinear.ErrorID);
	GroupData.Diag.sErrorText := 'MC_MoveLinearAbsolute error';
ELSIF fbGroupHalt.Error THEN
	GroupData.Diag.udiActualErrorID := TO_UDINT(fbGroupHalt.ErrorID);
	GroupData.Diag.sErrorText := 'MC_GroupHalt error';
ELSIF fbGroupStop.Error THEN
	GroupData.Diag.udiActualErrorID := TO_UDINT(fbGroupStop.ErrorID);
	GroupData.Diag.sErrorText := 'MC_GroupStop error';
ELSE
    GroupData.Diag.udiActualErrorID := UDINT#0;
    GroupData.Diag.sErrorText := '';
END_IF;

IF GroupData.Diag.udiActualErrorID <> UDINT#0 THEN
    GroupData.Diag.udiLastErrorID := GroupData.Diag.udiActualErrorID;
END_IF;

// Сохраняем последнюю ненулевую ошибку и формируем удобное представление для HMI.
IF (GroupData.Error.dwMotionErrorLatched <> DWORD#0)
OR (GroupData.Error.dwLogicalErrorLatched <> DWORD#0) THEN
	GroupData.Error.dwMotionErrorLast := GroupData.Error.dwMotionErrorLatched;
	GroupData.Error.dwLogicalErrorLast := GroupData.Error.dwLogicalErrorLatched;
END_IF;

GroupData.Error.stErrorActive := UpdateErrorView(
	dwMotionError := GroupData.Error.dwMotionErrorLatched OR GroupData.Error.dwMotionErrorActive,
	dwLogicalError := GroupData.Error.dwLogicalErrorLatched
);
GroupData.Error.stErrorLast := UpdateErrorView(
	dwMotionError := GroupData.Error.dwMotionErrorLast,
	dwLogicalError := GroupData.Error.dwLogicalErrorLast
);

// Для общей кнопки публикуется готовность владельца группы, а не только
// состояние диагностического инжектора.
FaultStatus.xResetAllowed := (GroupData.Diag.iStep = E_AXIS_GROUP_STATE.ERROR)
	AND xResetPermit
	AND NOT GroupData.Command.xGlobalError
	AND (GroupData.Status.xLocalError
		OR GroupData.Status.xLogicalError
		OR GroupData.Status.xGroupError);

METHOD UpdateErrorView : ST_AXIS_GROUP_ERROR
VAR_INPUT
	dwMotionError : DWORD; // Маска ошибок блоков SoftMotion
	dwLogicalError: DWORD; // Маска логических ошибок группы
END_VAR
VAR
	stError : ST_AXIS_GROUP_ERROR; // Представление ошибок отдельными флагами
END_VAR
stError.ENABLE_ERROR := (dwMotionError AND MOTION_ERR_ENABLE) <> DWORD#0;
// Зарезервировано для совместимости символов: питанием осей владеют FB_AXIS.
stError.POWER_ERROR := FALSE;
stError.DISABLE_ERROR := (dwMotionError AND MOTION_ERR_DISABLE) <> DWORD#0;
stError.RESET_ERROR := (dwMotionError AND MOTION_ERR_RESET) <> DWORD#0;
stError.MOVE_DIRECT_ERROR := (dwMotionError AND MOTION_ERR_MOVE_DIRECT) <> DWORD#0;
stError.MOVE_LINEAR_ERROR := (dwMotionError AND MOTION_ERR_MOVE_LINEAR) <> DWORD#0;
stError.HALT_ERROR := (dwMotionError AND MOTION_ERR_HALT) <> DWORD#0;
stError.STOP_ERROR := (dwMotionError AND MOTION_ERR_STOP) <> DWORD#0;
stError.READ_POSITION_ERROR := (dwMotionError AND MOTION_ERR_READ_POSITION) <> DWORD#0;
stError.READ_STATUS_ERROR := (dwMotionError AND MOTION_ERR_READ_STATUS) <> DWORD#0;
stError.READ_GROUP_ERROR := (dwMotionError AND MOTION_ERR_READ_GROUP_ERROR) <> DWORD#0;
stError.GROUP_ERROR_STOP := (dwMotionError AND MOTION_ERR_GROUP_ERROR_STOP) <> DWORD#0;
stError.SIMULATED_ERROR := (dwMotionError AND MOTION_ERR_SIMULATED) <> DWORD#0;
stError.OVERRIDE_ERROR := (dwMotionError AND MOTION_ERR_OVERRIDE) <> DWORD#0;

stError.STEP_TIMEOUT := (dwLogicalError AND LOG_STEP_TIMEOUT) <> DWORD#0;
stError.INVALID_STATE := (dwLogicalError AND LOG_INVALID_STATE) <> DWORD#0;
stError.POWER_PERMIT_READY := (dwLogicalError AND LOG_POWER_PERMIT_READY) <> DWORD#0;
stError.POWER_PERMIT_LOST := (dwLogicalError AND LOG_POWER_PERMIT_LOST_DIRECT) <> DWORD#0;

UpdateErrorView := stError;
END_METHOD

END_FUNCTION_BLOCK

// Device/Application/FB/FB_FAULT_INJECTOR/FB_AXIS_GROUP_FAULT_INJECTOR
FUNCTION_BLOCK FB_AXIS_GROUP_FAULT_INJECTOR
VAR_INPUT
	Request       : ST_AXIS_GROUP_FAULT_REQUEST; // Команда диагностической ошибки SM3
	xOwnerAllowed : BOOL; // Безопасные условия, рассчитанные FB_AXIS_GROUP
	xReset        : BOOL; // Штатный сброс группы
	Position      : SMC_POS_REF; // Текущая позиция для команды без перемещения
END_VAR
VAR_OUTPUT
	xError    : BOOL; // Защёлкнутая ошибка тестового Motion FB
	udiErrorID: UDINT; // ErrorID тестового Motion FB
	Status    : ST_FAULT_INJECTION_STATUS; // Состояние источника для HMI
END_VAR
VAR_IN_OUT
	AxisGroup : AXIS_GROUP_REF_SM3; // Ссылка на группу осей SoftMotion
END_VAR
VAR
	fbInvalidMove : MC_MoveDirectAbsolute; // Motion FB с недопустимым параметром
	rtExecute     : R_TRIG; // Фронт запроса HMI
	xExecute      : BOOL; // Execute удерживается до Error или Done
	xErrorLatched : BOOL; // Ошибка хранится до штатного сброса группы
END_VAR

rtExecute(CLK := Request.xExecute);

Status.xRejected := FALSE;
Status.xAllowed := Request.xEnabled AND xOwnerAllowed;

IF xReset THEN
	xExecute := FALSE;
	xErrorLatched := FALSE;
	udiErrorID := UDINT#0;
END_IF;

IF rtExecute.Q THEN
	IF Status.xAllowed THEN
		xExecute := TRUE;
	ELSE
		Status.xRejected := TRUE;
		Status.udiRejectSequence := Status.udiRejectSequence + UDINT#1;
		IF Status.udiRejectSequence = UDINT#0 THEN
			Status.udiRejectSequence := UDINT#1;
		END_IF;
	END_IF;
END_IF;

// По контракту SM3_Robotics VelFactor должен находиться в диапазоне ]0, 1].
// Отрицательное значение формирует Error/ErrorID без принятого перемещения.
fbInvalidMove(
	AxisGroup   := AxisGroup,
	Execute     := xExecute,
	Position    := Position,
	CoordSystem := SMC_COORD_SYSTEM.MCS,
	BufferMode  := MC_BUFFER_MODE.Aborting,
	VelFactor   := -1.0,
	AccFactor   := 1.0,
	JerkFactor  := 1.0
);

IF fbInvalidMove.Error THEN
	xErrorLatched := TRUE;
	udiErrorID := TO_UDINT(fbInvalidMove.ErrorID);
END_IF;

IF fbInvalidMove.Error OR fbInvalidMove.Done THEN
	xExecute := FALSE;
END_IF;

xError := xErrorLatched;
Status.xActive := xErrorLatched;
Status.xBusy := xExecute OR fbInvalidMove.Busy;
Status.xResetAllowed := xErrorLatched AND NOT Status.xBusy;

END_FUNCTION_BLOCK

// Device/Application/FB/FB_SIMULATION_DYNAMIC_LIMITS
FUNCTION_BLOCK FB_SIMULATION_DYNAMIC_LIMITS
VAR_INPUT
	xSimulationMode : BOOL; // Активна тестовая среда SIMULATION
	xSoftMotionMode : BOOL; // Роботом управляют локальные оси SoftMotion
	xAccelerationEnabled : BOOL; // Для следующего теста выбран ускоренный профиль
	xPrepareTest : BOOL; // Фронт подготовки следующего сценария
	uiRequestedFactor : UINT; // Запрошенное масштабирование времени 1..100
	xCellRunning : BOOL;
	xRobotBusy : BOOL;
	xMotionBusy : BOOL;
	xDrivesPowered : BOOL;
	xDrivesOff : BOOL;
	eGroupState : E_AXIS_GROUP_STATE;
	tTransactionTimeout : TIME := T#60S; // Общий предел Stop -> Disable -> Change -> Enable
END_VAR
VAR_OUTPUT
	xCellStopRequest : BOOL; // Сначала остановить технологический цикл
	xMotionStopRequest : BOOL; // Затем остановить движение группы
	xGroupDisableRequest : BOOL; // Перед изменением лимитов получить GroupDisabled
	xDrivesEnableRequest : BOOL; // После изменения вернуть штатную готовность
	xBusy : BOOL;
	xPending : BOOL; // Ползунок изменён; значение ждёт границы следующего теста
	xReadyForTest : BOOL; // Новый тест можно запускать
	xAccelerationActive : BOOL;
	uiAppliedFactor : UINT := UINT#1;
	xDone : BOOL;
	xError : BOOL;
	udiErrorId : UDINT;
END_VAR
VAR_IN_OUT
	AxisX : AXIS_REF_SM3;
	AxisY : AXIS_REF_SM3;
	AxisZ : AXIS_REF_SM3;
END_VAR
VAR CONSTANT
	STATE_IDLE : UINT := UINT#0;
	STATE_WAIT_STANDSTILL : UINT := UINT#10;
	STATE_WAIT_GROUP_DISABLED : UINT := UINT#20;
	STATE_CHANGE_X : UINT := UINT#30;
	STATE_CHANGE_Y : UINT := UINT#40;
	STATE_CHANGE_Z : UINT := UINT#50;
	STATE_PREPARE_ROLLBACK : UINT := UINT#55;
	STATE_WAIT_REENABLE : UINT := UINT#60;
	STATE_LOCKED_ERROR : UINT := UINT#90;
	ERR_INVALID_ORIGINAL_LIMITS : UDINT := UDINT#16#80010001;
	ERR_TRANSACTION_TIMEOUT : UDINT := UDINT#16#80010002;
	ERR_INVALID_STATE : UDINT := UDINT#16#80010003;
END_VAR
VAR
	rtPrepareTest : R_TRIG;
	tonTransaction : TON;
	uiState : UINT := UINT#0;
	uiAxis : UINT;
	uiDesiredFactor : UINT := UINT#1;
	uiTargetFactor : UINT := UINT#1;
	xOriginalLimitsSaved : BOOL;
	xOriginalLimitsValid : BOOL;
	xRestoreOnExit : BOOL;
	xRollback : BOOL;
	xReenableAfterChange : BOOL;

	alrOriginalVelocity : ARRAY [1..3] OF LREAL;
	alrOriginalAcceleration : ARRAY [1..3] OF LREAL;
	alrOriginalDeceleration : ARRAY [1..3] OF LREAL;
	alrOriginalJerk : ARRAY [1..3] OF LREAL;
	alrTargetVelocity : ARRAY [1..3] OF LREAL;
	alrTargetAcceleration : ARRAY [1..3] OF LREAL;
	alrTargetDeceleration : ARRAY [1..3] OF LREAL;
	alrTargetJerk : ARRAY [1..3] OF LREAL;
	lrFactor : LREAL;
	lrFactorSquared : LREAL;
	lrFactorCubed : LREAL;

	fbChangeX : SMC_ChangeDynamicLimits;
	fbChangeY : SMC_ChangeDynamicLimits;
	fbChangeZ : SMC_ChangeDynamicLimits;
END_VAR

// Запрошенное значение разрешено менять когда угодно. Оно только создаёт
// pending-запрос; уже выполняемая траектория никогда не перепланируется.
uiDesiredFactor := MAX(UINT#1, MIN(UINT#100, uiRequestedFactor));
IF NOT (xSimulationMode AND xSoftMotionMode AND xAccelerationEnabled) THEN
	uiDesiredFactor := UINT#1;
END_IF;
rtPrepareTest(CLK := xPrepareTest);

xCellStopRequest := FALSE;
xMotionStopRequest := FALSE;
xGroupDisableRequest := FALSE;
xDrivesEnableRequest := FALSE;
xDone := FALSE;

// Штатные лимиты снимаются ровно при входе в SoftMotion-симуляцию, до первого
// масштабирования. Прямое редактирование AXIS_REF здесь не выполняется.
IF xSimulationMode AND xSoftMotionMode AND NOT xOriginalLimitsSaved THEN
	// Dynamic limits из конфигуратора оси находятся в fSWMax*. fMax* — это
	// remote limits самого привода и у виртуальной оси законно остаются нулями.
	alrOriginalVelocity[1] := AxisX.fSWMaxVelocity;
	alrOriginalAcceleration[1] := AxisX.fSWMaxAcceleration;
	alrOriginalDeceleration[1] := AxisX.fSWMaxDeceleration;
	alrOriginalJerk[1] := AxisX.fSWMaxJerk;
	alrOriginalVelocity[2] := AxisY.fSWMaxVelocity;
	alrOriginalAcceleration[2] := AxisY.fSWMaxAcceleration;
	alrOriginalDeceleration[2] := AxisY.fSWMaxDeceleration;
	alrOriginalJerk[2] := AxisY.fSWMaxJerk;
	alrOriginalVelocity[3] := AxisZ.fSWMaxVelocity;
	alrOriginalAcceleration[3] := AxisZ.fSWMaxAcceleration;
	alrOriginalDeceleration[3] := AxisZ.fSWMaxDeceleration;
	alrOriginalJerk[3] := AxisZ.fSWMaxJerk;

	IF alrOriginalVelocity[1] <= LREAL#0.0 THEN alrOriginalVelocity[1] := AxisX.fMaxVelocity; END_IF;
	IF alrOriginalAcceleration[1] <= LREAL#0.0 THEN alrOriginalAcceleration[1] := AxisX.fMaxAcceleration; END_IF;
	IF alrOriginalDeceleration[1] <= LREAL#0.0 THEN alrOriginalDeceleration[1] := AxisX.fMaxDeceleration; END_IF;
	IF alrOriginalJerk[1] <= LREAL#0.0 THEN alrOriginalJerk[1] := AxisX.fMaxJerk; END_IF;
	IF alrOriginalVelocity[2] <= LREAL#0.0 THEN alrOriginalVelocity[2] := AxisY.fMaxVelocity; END_IF;
	IF alrOriginalAcceleration[2] <= LREAL#0.0 THEN alrOriginalAcceleration[2] := AxisY.fMaxAcceleration; END_IF;
	IF alrOriginalDeceleration[2] <= LREAL#0.0 THEN alrOriginalDeceleration[2] := AxisY.fMaxDeceleration; END_IF;
	IF alrOriginalJerk[2] <= LREAL#0.0 THEN alrOriginalJerk[2] := AxisY.fMaxJerk; END_IF;
	IF alrOriginalVelocity[3] <= LREAL#0.0 THEN alrOriginalVelocity[3] := AxisZ.fMaxVelocity; END_IF;
	IF alrOriginalAcceleration[3] <= LREAL#0.0 THEN alrOriginalAcceleration[3] := AxisZ.fMaxAcceleration; END_IF;
	IF alrOriginalDeceleration[3] <= LREAL#0.0 THEN alrOriginalDeceleration[3] := AxisZ.fMaxDeceleration; END_IF;
	IF alrOriginalJerk[3] <= LREAL#0.0 THEN alrOriginalJerk[3] := AxisZ.fMaxJerk; END_IF;

	xOriginalLimitsValid := TRUE;
	FOR uiAxis := UINT#1 TO UINT#3 DO
		xOriginalLimitsValid := xOriginalLimitsValid
			AND (alrOriginalVelocity[uiAxis] > LREAL#0.0)
			AND (alrOriginalAcceleration[uiAxis] > LREAL#0.0)
			AND (alrOriginalDeceleration[uiAxis] > LREAL#0.0)
			AND (alrOriginalJerk[uiAxis] > LREAL#0.0);
	END_FOR;
	IF xOriginalLimitsValid THEN
		xOriginalLimitsSaved := TRUE;
		uiAppliedFactor := UINT#1;
		xError := FALSE;
		udiErrorId := UDINT#0;
	ELSIF rtPrepareTest.Q THEN
		// До подготовки теста просто ждём инициализацию осей; не защёлкиваем
		// ложную ошибку на первом цикле после переключения среды.
		xError := TRUE;
		udiErrorId := ERR_INVALID_ORIGINAL_LIMITS;
	END_IF;
END_IF;

// Ошибка чтения исходных лимитов не должна блокировать обычную ячейку после
// выхода из тестовой среды и не должна переживать Online Change этого исправления.
IF NOT xSimulationMode
AND NOT xOriginalLimitsSaved
AND (uiState = STATE_IDLE)
AND (udiErrorId = ERR_INVALID_ORIGINAL_LIMITS) THEN
	xError := FALSE;
	udiErrorId := UDINT#0;
END_IF;

xRestoreOnExit := xOriginalLimitsSaved
	AND (NOT xSimulationMode OR NOT xSoftMotionMode)
	AND (uiAppliedFactor <> UINT#1);
xPending := xOriginalLimitsSaved AND (uiDesiredFactor <> uiAppliedFactor);

// Один общий таймаут защищает всю транзакцию Stop -> Disable -> Change -> Enable.
tonTransaction(IN := uiState <> STATE_IDLE, PT := tTransactionTimeout);
IF tonTransaction.Q
AND (uiState <> STATE_IDLE)
AND (uiState <> STATE_LOCKED_ERROR) THEN
	xError := TRUE;
	udiErrorId := ERR_TRANSACTION_TIMEOUT;
	uiState := STATE_LOCKED_ERROR;
END_IF;

CASE uiState OF
	STATE_IDLE:
		xBusy := FALSE;
		// Возврат штатных лимитов при выходе из SIMULATION выполняется сразу.
		// Обычная ячейка не получит Start, пока транзакция не закончена.
		IF xRestoreOnExit THEN
			xError := FALSE;
			udiErrorId := UDINT#0;
			uiTargetFactor := UINT#1;
			xRollback := FALSE;
			xReenableAfterChange := xSoftMotionMode AND NOT xDrivesOff;
			xBusy := TRUE;
			uiState := STATE_WAIT_STANDSTILL;
		ELSIF rtPrepareTest.Q
		AND xSimulationMode
		AND xSoftMotionMode
		AND xPending
		AND NOT xCellRunning THEN
			xError := FALSE;
			udiErrorId := UDINT#0;
			uiTargetFactor := uiDesiredFactor;
			xRollback := FALSE;
			xReenableAfterChange := NOT xDrivesOff;
			xBusy := TRUE;
			uiState := STATE_WAIT_STANDSTILL;
		ELSIF NOT xSimulationMode
		AND xOriginalLimitsSaved
		AND (uiAppliedFactor = UINT#1) THEN
			// Лимиты не менялись либо уже успешно восстановлены.
			xOriginalLimitsSaved := FALSE;
		END_IF;

	STATE_WAIT_STANDSTILL:
		xBusy := TRUE;
		xCellStopRequest := xCellRunning;
		xMotionStopRequest := xMotionBusy OR xRobotBusy;
		IF NOT xCellRunning AND NOT xMotionBusy AND NOT xRobotBusy THEN
			uiState := STATE_WAIT_GROUP_DISABLED;
		END_IF;

	STATE_WAIT_GROUP_DISABLED:
		xBusy := TRUE;
		xGroupDisableRequest := NOT xDrivesOff;
		IF xDrivesOff AND (eGroupState = E_AXIS_GROUP_STATE.DISABLED) THEN
			IF xRollback THEN
				FOR uiAxis := UINT#1 TO UINT#3 DO
					alrTargetVelocity[uiAxis] := alrOriginalVelocity[uiAxis];
					alrTargetAcceleration[uiAxis] := alrOriginalAcceleration[uiAxis];
					alrTargetDeceleration[uiAxis] := alrOriginalDeceleration[uiAxis];
					alrTargetJerk[uiAxis] := alrOriginalJerk[uiAxis];
				END_FOR;
			ELSE
				lrFactor := UINT_TO_LREAL(uiTargetFactor);
				lrFactorSquared := lrFactor * lrFactor;
				lrFactorCubed := lrFactorSquared * lrFactor;
				alrTargetVelocity[1] := alrOriginalVelocity[1] * lrFactor;
				alrTargetAcceleration[1] := alrOriginalAcceleration[1] * lrFactorSquared;
				alrTargetDeceleration[1] := alrOriginalDeceleration[1] * lrFactorSquared;
				alrTargetJerk[1] := alrOriginalJerk[1] * lrFactorCubed;
				alrTargetVelocity[2] := alrOriginalVelocity[2] * lrFactor;
				alrTargetAcceleration[2] := alrOriginalAcceleration[2] * lrFactorSquared;
				alrTargetDeceleration[2] := alrOriginalDeceleration[2] * lrFactorSquared;
				alrTargetJerk[2] := alrOriginalJerk[2] * lrFactorCubed;
				alrTargetVelocity[3] := alrOriginalVelocity[3] * lrFactor;
				alrTargetAcceleration[3] := alrOriginalAcceleration[3] * lrFactorSquared;
				alrTargetDeceleration[3] := alrOriginalDeceleration[3] * lrFactorSquared;
				alrTargetJerk[3] := alrOriginalJerk[3] * lrFactorCubed;
			END_IF;
			uiState := STATE_CHANGE_X;
		END_IF;

	STATE_CHANGE_X:
		xBusy := TRUE;
		IF fbChangeX.bError THEN
			xError := TRUE;
			udiErrorId := TO_UDINT(fbChangeX.ErrorID);
			IF xRollback THEN uiState := STATE_LOCKED_ERROR;
			ELSE uiState := STATE_PREPARE_ROLLBACK; END_IF;
		ELSIF fbChangeX.bDone THEN
			uiState := STATE_CHANGE_Y;
		END_IF;

	STATE_CHANGE_Y:
		xBusy := TRUE;
		IF fbChangeY.bError THEN
			xError := TRUE;
			udiErrorId := TO_UDINT(fbChangeY.ErrorID);
			IF xRollback THEN uiState := STATE_LOCKED_ERROR;
			ELSE uiState := STATE_PREPARE_ROLLBACK; END_IF;
		ELSIF fbChangeY.bDone THEN
			uiState := STATE_CHANGE_Z;
		END_IF;

	STATE_CHANGE_Z:
		xBusy := TRUE;
		IF fbChangeZ.bError THEN
			xError := TRUE;
			udiErrorId := TO_UDINT(fbChangeZ.ErrorID);
			IF xRollback THEN uiState := STATE_LOCKED_ERROR;
			ELSE uiState := STATE_PREPARE_ROLLBACK; END_IF;
		ELSIF fbChangeZ.bDone THEN
			IF xReenableAfterChange THEN
				uiState := STATE_WAIT_REENABLE;
			ELSE
				IF xRollback THEN uiAppliedFactor := UINT#1;
				ELSE uiAppliedFactor := uiTargetFactor; END_IF;
				xDone := NOT xRollback;
				xBusy := FALSE;
				uiState := STATE_IDLE;
			END_IF;
		END_IF;

	STATE_PREPARE_ROLLBACK:
		// Один цикл с Execute=FALSE создаёт корректный новый фронт для X.
		xBusy := TRUE;
		xRollback := TRUE;
		uiState := STATE_WAIT_GROUP_DISABLED;

	STATE_WAIT_REENABLE:
		xBusy := TRUE;
		xDrivesEnableRequest := TRUE;
		IF xDrivesPowered AND (eGroupState = E_AXIS_GROUP_STATE.READY) THEN
			IF xRollback THEN uiAppliedFactor := UINT#1;
			ELSE uiAppliedFactor := uiTargetFactor; END_IF;
			xDone := NOT xRollback;
			xBusy := FALSE;
			uiState := STATE_IDLE;
		END_IF;

	STATE_LOCKED_ERROR:
		// При неизвестном/неустранимом результате оставляем группу отключённой.
		// Следующий Start заблокирован, пока инженер не устранит причину.
		xBusy := FALSE;
		xGroupDisableRequest := NOT xDrivesOff;

ELSE
	xError := TRUE;
	udiErrorId := ERR_INVALID_STATE;
	uiState := STATE_LOCKED_ERROR;
END_CASE;

fbChangeX(
	Axis := AxisX,
	bExecute := uiState = STATE_CHANGE_X,
	fMaxVelocity := alrTargetVelocity[1],
	fMaxAcceleration := alrTargetAcceleration[1],
	fMaxDeceleration := alrTargetDeceleration[1],
	fMaxJerk := alrTargetJerk[1]
);
fbChangeY(
	Axis := AxisY,
	bExecute := uiState = STATE_CHANGE_Y,
	fMaxVelocity := alrTargetVelocity[2],
	fMaxAcceleration := alrTargetAcceleration[2],
	fMaxDeceleration := alrTargetDeceleration[2],
	fMaxJerk := alrTargetJerk[2]
);
fbChangeZ(
	Axis := AxisZ,
	bExecute := uiState = STATE_CHANGE_Z,
	fMaxVelocity := alrTargetVelocity[3],
	fMaxAcceleration := alrTargetAcceleration[3],
	fMaxDeceleration := alrTargetDeceleration[3],
	fMaxJerk := alrTargetJerk[3]
);

xPending := xOriginalLimitsSaved AND (uiDesiredFactor <> uiAppliedFactor);
xAccelerationActive := xSimulationMode AND xSoftMotionMode
	AND (uiAppliedFactor > UINT#1) AND NOT xError;
xReadyForTest := NOT xBusy AND NOT xError
	AND (NOT (xSimulationMode AND xSoftMotionMode AND xAccelerationEnabled) OR NOT xPending);

END_FUNCTION_BLOCK

// Device/Application/FB/FB_MOTION_MANAGER
FUNCTION_BLOCK FB_MOTION_MANAGER
VAR_INPUT
	stPoint : ARRAY [0..GVL_POINT.iPointNumber] OF ST_POINT; // Глобальная таблица точек
	xReset  : BOOL; // Сброс ошибок менеджера движения
	FaultRequest : ST_POINT_FAULT_REQUEST; // Диагностические ошибки проверки точки
	xSpeedFactorOverride : BOOL; // Для отдельной проверки точки с телефона
	lrSpeedFactorOverride : LREAL; // 0.001..1.0, применяется вместо SpeedFactor точки
	lrAccelerationFactor : LREAL := 1.0; // Единый предел разгона/торможения группы 0.01..1.0
	lrJerkFactor : LREAL := 1.0; // Плавность групповой траектории 0.01..1.0
END_VAR
VAR_OUTPUT
	FaultStatus : ST_FAULT_INJECTION_STATUS; // Состояние инжектора проверки точки
END_VAR
VAR
	curPoint      : ST_POINT; // Координаты выбранной точки
	curPointName  : E_POINT_NAME; // Имя выбранной точки
	fbPointManager: FB_POINT_MANAGER; // Проверка координат и скорости точки
	fbPointFaultInjector : FB_POINT_FAULT_INJECTOR; // Безопасная подмена проверяемой точки
	rtReset       : R_TRIG; // Фронт команды сброса менеджера движения
	xFaultAllowed : BOOL; // Менеджер готов к синтетической проверке без движения
	xGroupMotionStarted : BOOL; // Группа приняла движение, ожидание запуска завершено
	tonMotionStart : TON; // Общий предел проверки точки и старта группы
END_VAR
VAR CONSTANT
	ERR_POINT_INVALID : DWORD := DWORD#16#0000_0001; // Недопустимая точка
	ERR_GROUP         : DWORD := DWORD#16#0000_0002; // Ошибка группы осей
	ERR_GLOBAL_STOP   : DWORD := DWORD#16#0000_0004; // Глобальная ошибка ячейки
	ERR_START_TIMEOUT : DWORD := DWORD#16#0000_0008; // Проверка/запуск группы не завершены вовремя
	WRN_RESET_GLOBAL_ERROR : UINT := 1; // Глобальная ошибка ещё активна
	WRN_SIM_ERROR_NOT_ALLOWED : UINT := 2; // Тестовая проверка запрещена текущим состоянием
END_VAR
VAR_IN_OUT
	stMotionManager : ST_MOTION_MANAGER; // Команды, статусы и диагностика менеджера движения
	GroupData       : ST_AXIS_GROUP; // Команды, статусы и диагностика группы XYZ
	stPointManager  : ST_POINT_MANAGER; // Команды, статусы и диагностика проверки точки
END_VAR

xFaultAllowed := (stMotionManager.Diag.eState = E_MOTION_MANAGER_STATE.IDLE)
	AND NOT stMotionManager.Command.xExecute
	AND NOT stMotionManager.Command.xGlobalError
	AND (stMotionManager.Error.dwErrorActive = DWORD#0)
	AND NOT GroupData.Status.xLocalError
	AND NOT GroupData.Command.xMoveDirect
	AND NOT GroupData.Command.xMoveLinear;

fbPointFaultInjector(
	Request := FaultRequest,
	xOwnerAllowed := xFaultAllowed,
	xComplete := stMotionManager.Diag.eState = E_MOTION_MANAGER_STATE.ERROR,
	PointRaw := stPoint[E_POINT_NAME.MAGAZINE_DETAIL]
);
FaultStatus := fbPointFaultInjector.Status;

IF fbPointFaultInjector.Status.xRejected THEN
	stPointManager.Diag.stWarning.uiCode := WRN_SIM_ERROR_NOT_ALLOWED;
	stPointManager.Diag.stWarning.udiSequence := stPointManager.Diag.stWarning.udiSequence + UDINT#1;
	IF stPointManager.Diag.stWarning.udiSequence = UDINT#0 THEN
		stPointManager.Diag.stWarning.udiSequence := UDINT#1;
	END_IF;
END_IF;

IF fbPointFaultInjector.xExecute THEN
	curPoint := fbPointFaultInjector.Point;
	curPointName := E_POINT_NAME.NONE;
END_IF;

// Рабочая точка должна быть защёлкнута до вызова FB_POINT_MANAGER. Иначе при
// переходе в VALIDATE менеджер точек видит curPoint от предыдущей команды
// (или нулевой ST_POINT при первом проходе), потому что прежняя запись
// выполнялась ниже вызова FB_POINT_MANAGER в CASE VALIDATE.
IF (stMotionManager.Diag.eState = E_MOTION_MANAGER_STATE.VALIDATE)
AND NOT fbPointFaultInjector.xExecute THEN

	curPoint := stPoint[stMotionManager.Command.eTargetPoint];
	curPointName := stMotionManager.Command.eTargetPoint;
END_IF;

fbPointManager(
			stPointManager := stPointManager,
			stPoint := curPoint
		);
		
stMotionManager.Status.xBusy := FALSE;
stMotionManager.Status.xDone := FALSE;
stMotionManager.Status.xError := FALSE;
stMotionManager.Status.xReady:= FALSE;
stMotionManager.Command.xReset := xReset;
rtReset(CLK := xReset);

IF rtReset.Q
AND (stMotionManager.Diag.eState = E_MOTION_MANAGER_STATE.ERROR)
AND stMotionManager.Command.xGlobalError THEN
	stMotionManager.Diag.stWarning.uiCode := WRN_RESET_GLOBAL_ERROR;
	stMotionManager.Diag.stWarning.udiSequence := stMotionManager.Diag.stWarning.udiSequence + UDINT#1;
	IF stMotionManager.Diag.stWarning.udiSequence = UDINT#0 THEN
		stMotionManager.Diag.stWarning.udiSequence := UDINT#1;
	END_IF;
END_IF;


IF (stMotionManager.Diag.eState = E_MOTION_MANAGER_STATE.MOTION_SIM)
AND ((GroupData.Diag.iStep = E_AXIS_GROUP_STATE.MOVING_DIRECT)
	OR (GroupData.Status.xMoveDirectDone AND GroupData.Command.xMoveDirect)) THEN
	xGroupMotionStarted := TRUE;
END_IF;
tonMotionStart(
	IN := (stMotionManager.Diag.eState = E_MOTION_MANAGER_STATE.VALIDATE)
		OR ((stMotionManager.Diag.eState = E_MOTION_MANAGER_STATE.MOTION_SIM)
			AND NOT xGroupMotionStarted),
	PT := GroupData.Timeouts.tGroupTimeout
);

// Stop должен отменять ещё не запущенную команду и завершённую команду,
// ожидающую освобождения. Проверка точки тоже получает спад Execute.
IF stMotionManager.Command.xGlobalError THEN
	stPointManager.Command.xExecute := FALSE;
	GroupData.Command.xMoveDirect := FALSE;
	GroupData.Command.xMoveLinear := FALSE;
	stMotionManager.Error.dwErrorActive := stMotionManager.Error.dwErrorActive OR ERR_GLOBAL_STOP;
	stMotionManager.Diag.eState := E_MOTION_MANAGER_STATE.ERROR;
ELSIF stMotionManager.Command.xStop
AND (stMotionManager.Diag.eState <> E_MOTION_MANAGER_STATE.ERROR) THEN
	stPointManager.Command.xExecute := FALSE;
	GroupData.Command.xMoveDirect := FALSE;
	GroupData.Command.xMoveLinear := FALSE;
	xGroupMotionStarted := FALSE;
	stMotionManager.Diag.eState := E_MOTION_MANAGER_STATE.IDLE;
ELSIF tonMotionStart.Q THEN
	stPointManager.Command.xExecute := FALSE;
	GroupData.Command.xMoveDirect := FALSE;
	GroupData.Command.xMoveLinear := FALSE;
	stMotionManager.Error.dwErrorActive := stMotionManager.Error.dwErrorActive OR ERR_START_TIMEOUT;
	stMotionManager.Diag.eState := E_MOTION_MANAGER_STATE.ERROR;
END_IF;

CASE stMotionManager.Diag.eState OF 
	// --------------------------------------------------
	E_MOTION_MANAGER_STATE.IDLE:
	// --------------------------------------------------
		// Менеджер является единственным владельцем команд движения группы.
		// После завершения или сброса не оставляем уровень Execute защёлкнутым.
		GroupData.Command.xMoveDirect := FALSE;
		GroupData.Command.xMoveLinear := FALSE;
		xGroupMotionStarted := FALSE;
		stMotionManager.Status.xReady:= TRUE;
		IF (stMotionManager.Command.xExecute OR fbPointFaultInjector.xExecute)
		AND NOT stMotionManager.Command.xGlobalError
		AND NOT stMotionManager.Command.xStop THEN
			stMotionManager.Status.xBusy := TRUE;
			stMotionManager.Diag.eState := E_MOTION_MANAGER_STATE.VALIDATE;
		ELSIF stMotionManager.Command.xGlobalError THEN
			stMotionManager.Error.dwErrorActive := stMotionManager.Error.dwErrorActive OR ERR_GLOBAL_STOP;
			stMotionManager.Diag.eState := E_MOTION_MANAGER_STATE.ERROR;
		END_IF;
	
	// --------------------------------------------------
	E_MOTION_MANAGER_STATE.VALIDATE:
	// --------------------------------------------------
		stMotionManager.Status.xBusy := TRUE;
		stPointManager.Command.xExecute := TRUE;
		
		IF stPointManager.Status.xDone AND NOT stPointManager.Status.xInvalid THEN
			stPointManager.Command.xExecute := FALSE;
			IF stMotionManager.Command.xMode THEN
				stMotionManager.Diag.eState := 	E_MOTION_MANAGER_STATE.MOTION_MODBUS;
			ELSE
				stMotionManager.Diag.eState := 	E_MOTION_MANAGER_STATE.MOTION_SIM;
			END_IF;
		ELSIF stPointManager.Status.xDone AND stPointManager.Status.xInvalid THEN
			stPointManager.Command.xExecute := FALSE;
			stMotionManager.Error.dwErrorActive := stMotionManager.Error.dwErrorActive OR ERR_POINT_INVALID;
			stMotionManager.Diag.eState := 	E_MOTION_MANAGER_STATE.ERROR;
		END_IF;
	
	// --------------------------------------------------
	E_MOTION_MANAGER_STATE.MOTION_SIM:
	// --------------------------------------------------
	
		stMotionManager.Status.xBusy := TRUE;
		 
		GroupData.MotionParam.lrX := curPoint.X;
		GroupData.MotionParam.lrY := curPoint.Y;
		GroupData.MotionParam.lrZ := curPoint.Z;
		IF xSpeedFactorOverride THEN
			GroupData.MotionParam.VelFactor := LIMIT(0.001, lrSpeedFactorOverride, 1.0);
		ELSE
			GroupData.MotionParam.VelFactor := curPoint.SpeedFactor;
		END_IF;
		// У группы SoftMotion один AccFactor для обеих сторон профиля. PLC передаёт
		// сюда более строгий из глобальных процентов разгона и торможения.
		GroupData.MotionParam.AccFactor := LIMIT(0.01, lrAccelerationFactor, 1.0);
		GroupData.MotionParam.JerkFactor := LIMIT(0.01, lrJerkFactor, 1.0);
		IF GroupData.Diag.iStep = E_AXIS_GROUP_STATE.READY
		AND NOT GroupData.Command.xMoveDirect
		AND NOT stMotionManager.Command.xGlobalError
		AND NOT stMotionManager.Command.xStop THEN
			GroupData.Command.xMoveDirect := TRUE;
		END_IF;
		
		IF stMotionManager.Command.xStop THEN
			GroupData.Command.xMoveDirect := FALSE;
			GroupData.Command.xMoveLinear := FALSE;
			stMotionManager.Status.xBusy := FALSE;
			stMotionManager.Diag.eState := E_MOTION_MANAGER_STATE.IDLE;
		ELSIF GroupData.Status.xMoveDirectDone AND GroupData.Command.xMoveDirect THEN
			GroupData.Command.xMoveDirect := FALSE;
			stMotionManager.Status.eCurrentPoint := curPointName;
			stMotionManager.Diag.eState := 	E_MOTION_MANAGER_STATE.DONE;
		ELSIF GroupData.Diag.iStep = E_AXIS_GROUP_STATE.ERROR OR stMotionManager.Command.xGlobalError  THEN
			GroupData.Command.xMoveDirect := FALSE;
			GroupData.Command.xMoveLinear := FALSE;
			IF GroupData.Diag.iStep = E_AXIS_GROUP_STATE.ERROR THEN
				stMotionManager.Error.dwErrorActive := stMotionManager.Error.dwErrorActive OR ERR_GROUP;
			END_IF;
			IF stMotionManager.Command.xGlobalError THEN
				stMotionManager.Error.dwErrorActive := stMotionManager.Error.dwErrorActive OR ERR_GLOBAL_STOP;
			END_IF;
			stMotionManager.Diag.eState := 	E_MOTION_MANAGER_STATE.ERROR;
		END_IF;
	
	// --------------------------------------------------
	E_MOTION_MANAGER_STATE.ERROR:
	// --------------------------------------------------
		GroupData.Command.xMoveDirect := FALSE;
		GroupData.Command.xMoveLinear := FALSE;
		stMotionManager.Status.xError := TRUE;
		IF NOT stMotionManager.Command.xGlobalError AND stMotionManager.Command.xReset THEN
			stMotionManager.Error.dwErrorLast := stMotionManager.Error.dwErrorActive;
			stMotionManager.Error.dwErrorActive := DWORD#0;
			stMotionManager.Status.xError := FALSE;
			stMotionManager.Diag.eState := 	E_MOTION_MANAGER_STATE.IDLE;
		END_IF;
	
	
	// --------------------------------------------------
	E_MOTION_MANAGER_STATE.DONE:
	// --------------------------------------------------
		stMotionManager.Status.xBusy := FALSE;
		stMotionManager.Status.xDone := TRUE;
		IF NOT stMotionManager.Command.xExecute THEN
			stMotionManager.Diag.eState := 	E_MOTION_MANAGER_STATE.IDLE;
		END_IF;
	END_CASE;

// Журнал отражает состояние каждого FB, включая каскадные ошибки зависимостей.
stMotionManager.Error.dwAlarmActive := stMotionManager.Error.dwErrorActive;

stMotionManager.Error.stErrorActive := UpdateErrorView(
	dwError := stMotionManager.Error.dwErrorActive
);
stMotionManager.Error.stErrorLast := UpdateErrorView(
	dwError := stMotionManager.Error.dwErrorLast
);
FaultStatus.xResetAllowed := stMotionManager.Status.xError
	AND NOT FaultStatus.xBusy;

METHOD UpdateErrorView : ST_MOTION_MANAGER_ERROR
VAR_INPUT
	dwError : DWORD; // Битовая маска для расшифровки
END_VAR
VAR
	stError : ST_MOTION_MANAGER_ERROR; // Представление ошибок отдельными флагами
END_VAR
stError.POINT_INVALID := (dwError AND ERR_POINT_INVALID) <> DWORD#0;
stError.GROUP_ERROR := (dwError AND ERR_GROUP) <> DWORD#0;
stError.GLOBAL_STOP := (dwError AND ERR_GLOBAL_STOP) <> DWORD#0;
stError.START_TIMEOUT := (dwError AND ERR_START_TIMEOUT) <> DWORD#0;

UpdateErrorView := stError;
END_METHOD

END_FUNCTION_BLOCK

// Device/Application/FB/FB_POINT_MANAGER
FUNCTION_BLOCK FB_POINT_MANAGER
VAR_INPUT
	stPoint : ST_POINT; // Проверяемая точка
END_VAR
VAR_OUTPUT
END_VAR
VAR
END_VAR
VAR_IN_OUT
	stPointManager : ST_POINT_MANAGER; // Команды, статусы и диагностика проверки точки
END_VAR
VAR CONSTANT
	X_OUT_OF_LIMIT : DWORD := 1; // Координата X вне допустимых границ
	Y_OUT_OF_LIMIT : DWORD := 2; // Координата Y вне допустимых границ
	Z_OUT_OF_LIMIT : DWORD := 4; // Координата Z вне допустимых границ
	INVALID_VEL    : DWORD := 8; // Недопустимый коэффициент скорости
	X_LIMIT_CONFIG_INVALID : DWORD := 16; // Software limits оси X недоступны или некорректны
	Y_LIMIT_CONFIG_INVALID : DWORD := 32; // Software limits оси Y недоступны или некорректны
	Z_LIMIT_CONFIG_INVALID : DWORD := 64; // Software limits оси Z недоступны или некорректны
	POINT_NOT_CONFIGURED : DWORD := 128; // Инженерная точка не подтверждена редактором
END_VAR

stPointManager.Status.xBusy := FALSE;
stPointManager.Status.xDone := FALSE;
stPointManager.Status.xInvalid := FALSE;




CASE stPointManager.Diag.eState OF
	// --------------------------------------------------
	E_POINT_MANAGER_STATE.IDLE:
	// --------------------------------------------------
		stPointManager.Error.dwErrorActive := DWORD#0;
		IF stPointManager.Command.xExecute THEN
			stPointManager.Status.xBusy := TRUE;
			stPointManager.Diag.eState := E_POINT_MANAGER_STATE.CHECK_ZONE;
		END_IF

	// --------------------------------------------------
	E_POINT_MANAGER_STATE.CHECK_ZONE:
	// --------------------------------------------------
		stPointManager.Status.xBusy := TRUE;
		IF NOT stPoint.xConfigured THEN
			stPointManager.Error.dwErrorActive :=
				stPointManager.Error.dwErrorActive OR POINT_NOT_CONFIGURED;
		END_IF

		IF NOT stPointManager.Diag.xXLimitValid
		OR NOT stPointManager.Diag.xYLimitValid
		OR NOT stPointManager.Diag.xZLimitValid THEN
			// Без достоверных активных SoftMotion limits движение к точке запрещается.
			// Статический резервный диапазон здесь намеренно не применяется.
			IF NOT stPointManager.Diag.xXLimitValid THEN
				stPointManager.Error.dwErrorActive :=
					stPointManager.Error.dwErrorActive OR X_LIMIT_CONFIG_INVALID;
			END_IF
			IF NOT stPointManager.Diag.xYLimitValid THEN
				stPointManager.Error.dwErrorActive :=
					stPointManager.Error.dwErrorActive OR Y_LIMIT_CONFIG_INVALID;
			END_IF
			IF NOT stPointManager.Diag.xZLimitValid THEN
				stPointManager.Error.dwErrorActive :=
					stPointManager.Error.dwErrorActive OR Z_LIMIT_CONFIG_INVALID;
			END_IF
		ELSE
			IF NOT ((stPointManager.Diag.lrX_MinLimit <= stPoint.X) AND (stPoint.X <= stPointManager.Diag.lrX_MaxLimit)) THEN
				stPointManager.Error.dwErrorActive := stPointManager.Error.dwErrorActive OR X_OUT_OF_LIMIT;
			END_IF

			IF NOT ((stPointManager.Diag.lrY_MinLimit <= stPoint.Y) AND (stPoint.Y <= stPointManager.Diag.lrY_MaxLimit)) THEN
				stPointManager.Error.dwErrorActive := stPointManager.Error.dwErrorActive OR Y_OUT_OF_LIMIT;
			END_IF

			IF NOT ((stPointManager.Diag.lrZ_MinLimit <= stPoint.Z) AND (stPoint.Z <= stPointManager.Diag.lrZ_MaxLimit)) THEN
				stPointManager.Error.dwErrorActive := stPointManager.Error.dwErrorActive OR Z_OUT_OF_LIMIT;
			END_IF
		END_IF

		stPointManager.Diag.eState := E_POINT_MANAGER_STATE.CHECK_VEL_FACTOR;

	// --------------------------------------------------
	E_POINT_MANAGER_STATE.CHECK_VEL_FACTOR:
	// --------------------------------------------------
		stPointManager.Status.xBusy := TRUE;

		IF  NOT ((0.1 < stPoint.SpeedFactor) AND(stPoint.SpeedFactor <= 1.0))  THEN
			stPointManager.Error.dwErrorActive := stPointManager.Error.dwErrorActive OR INVALID_VEL;
		END_IF

		stPointManager.Diag.eState := E_POINT_MANAGER_STATE.CHECK_ALL;

	// --------------------------------------------------
	E_POINT_MANAGER_STATE.CHECK_ALL:
	// --------------------------------------------------
		stPointManager.Status.xDone := TRUE;
		stPointManager.Status.xBusy := FALSE;
		IF stPointManager.Error.dwErrorActive <> DWORD#0 THEN
			stPointManager.Status.xInvalid := TRUE;
			stPointManager.Error.dwErrorLast := stPointManager.Error.dwErrorActive;
		ELSE
			stPointManager.Status.xInvalid := FALSE;
		END_IF

		IF NOT stPointManager.Command.xExecute THEN
			stPointManager.Diag.eState := E_POINT_MANAGER_STATE.IDLE;
		END_IF

END_CASE

stPointManager.Error.dwAlarmActive := stPointManager.Error.dwErrorActive;

stPointManager.Error.stErrorActive := UpdateErrorView(
	dwError := stPointManager.Error.dwErrorActive
);
stPointManager.Error.stErrorLast := UpdateErrorView(
	dwError := stPointManager.Error.dwErrorLast
);

METHOD UpdateErrorView : ST_POINT_MANAGER_ERROR
VAR_INPUT
	dwError : DWORD; // Битовая маска для расшифровки
END_VAR
VAR
	stError : ST_POINT_MANAGER_ERROR; // Представление ошибок отдельными флагами
END_VAR
stError.X_OUT_OF_LIMIT := (dwError AND X_OUT_OF_LIMIT) <> DWORD#0;
stError.Y_OUT_OF_LIMIT := (dwError AND Y_OUT_OF_LIMIT) <> DWORD#0;
stError.Z_OUT_OF_LIMIT := (dwError AND Z_OUT_OF_LIMIT) <> DWORD#0;
stError.INVALID_VEL := (dwError AND INVALID_VEL) <> DWORD#0;
stError.X_LIMIT_CONFIG_INVALID := (dwError AND X_LIMIT_CONFIG_INVALID) <> DWORD#0;
stError.Y_LIMIT_CONFIG_INVALID := (dwError AND Y_LIMIT_CONFIG_INVALID) <> DWORD#0;
stError.Z_LIMIT_CONFIG_INVALID := (dwError AND Z_LIMIT_CONFIG_INVALID) <> DWORD#0;
stError.POINT_NOT_CONFIGURED := (dwError AND POINT_NOT_CONFIGURED) <> DWORD#0;

UpdateErrorView := stError;
END_METHOD

END_FUNCTION_BLOCK

// Device/Application/FB/FB_FAULT_INJECTOR/FB_POINT_FAULT_INJECTOR
FUNCTION_BLOCK FB_POINT_FAULT_INJECTOR
VAR_INPUT
	Request       : ST_POINT_FAULT_REQUEST; // Запросы конкретных ошибок точки
	xOwnerAllowed : BOOL; // Безопасные условия, рассчитанные менеджером движения
	xComplete     : BOOL; // Штатная ошибка уже сформирована владельцем
	PointRaw      : ST_POINT; // Исходная корректная точка
END_VAR
VAR_OUTPUT
	Point    : ST_POINT; // Точка, передаваемая штатной проверке
	xExecute : BOOL; // Синтетический запрос проверки без запуска движения
	Status   : ST_FAULT_INJECTION_STATUS; // Состояние источника для HMI
END_VAR
VAR
	rtXOutOfLimit     : R_TRIG;
	rtYOutOfLimit     : R_TRIG;
	rtZOutOfLimit     : R_TRIG;
	rtInvalidVelocity : R_TRIG;
	xRequestPulse     : BOOL;
	xInjectX          : BOOL;
	xInjectY          : BOOL;
	xInjectZ          : BOOL;
	xInjectVelocity   : BOOL;
END_VAR
VAR CONSTANT
	INVALID_COORDINATE : LREAL := 1.0E+09; // Заведомо вне рабочей зоны проверки
END_VAR

rtXOutOfLimit(CLK := Request.xXOutOfLimit);
rtYOutOfLimit(CLK := Request.xYOutOfLimit);
rtZOutOfLimit(CLK := Request.xZOutOfLimit);
rtInvalidVelocity(CLK := Request.xInvalidVelocity);

xRequestPulse := rtXOutOfLimit.Q
	OR rtYOutOfLimit.Q
	OR rtZOutOfLimit.Q
	OR rtInvalidVelocity.Q;

Status.xRejected := FALSE;
Status.xAllowed := Request.xEnabled AND xOwnerAllowed;

IF xComplete THEN
	xInjectX := FALSE;
	xInjectY := FALSE;
	xInjectZ := FALSE;
	xInjectVelocity := FALSE;
END_IF;

IF xRequestPulse THEN
	IF Status.xAllowed THEN
		xInjectX := rtXOutOfLimit.Q;
		xInjectY := rtYOutOfLimit.Q;
		xInjectZ := rtZOutOfLimit.Q;
		xInjectVelocity := rtInvalidVelocity.Q;
	ELSE
		Status.xRejected := TRUE;
		Status.udiRejectSequence := Status.udiRejectSequence + UDINT#1;
		IF Status.udiRejectSequence = UDINT#0 THEN
			Status.udiRejectSequence := UDINT#1;
		END_IF;
	END_IF;
END_IF;

Point := PointRaw;
// Диагностическая инъекция проверяет выбранный дефект, а не состояние
// инженерного хранилища точек.
IF xInjectX OR xInjectY OR xInjectZ OR xInjectVelocity THEN
	Point.xConfigured := TRUE;
END_IF;
IF xInjectX THEN
	Point.X := INVALID_COORDINATE;
END_IF;
IF xInjectY THEN
	Point.Y := INVALID_COORDINATE;
END_IF;
IF xInjectZ THEN
	Point.Z := INVALID_COORDINATE;
END_IF;
IF xInjectVelocity THEN
	Point.SpeedFactor := 0.0;
END_IF;

xExecute := xInjectX OR xInjectY OR xInjectZ OR xInjectVelocity;
Status.xActive := xExecute;
Status.xBusy := xExecute;
Status.xResetAllowed := FALSE;

END_FUNCTION_BLOCK

// Device/Application/FB/FB_MACHINE
FUNCTION_BLOCK FB_MACHINE
VAR_INPUT
	xIoManual : BOOL; // Прямое ручное I/O отменяет рецепт и сохраняет аварии
	xTestInitialize : BOOL;
	uiTestInitialState : UINT;
	uiTestProductType : UINT;
	xExecute          : BOOL; // Запуск разрешённой операции обслуживания
    xReset            : BOOL; // Сброс ошибки конкретного станка
	xResetGlobal      : BOOL; // Общий сброс ошибок ячейки
	xGlobalError      : BOOL; // Глобальная ошибка ячейки
	xManualMode       : BOOL; // Ручной режим: открытая операторская дверь не формирует аварию обслуживания
	xAutomaticUseEnabled : BOOL; // Станок выбран для автоматической обработки
	xPointsConfigured : BOOL; // Настроены ABOVE, CHUCK_APROACH и CHUCK_POSITION этого станка
	xRobotMotionBusy   : BOOL; // Группа/ось робота ещё движется или тормозит
	xSafetyDoorControlEnabled : BOOL := TRUE; // Модель двери; FALSE для ручной двери в NORMAL
	xHmiOpenSafetyDoor  : BOOL; // Импульс ручного открытия операторской двери
	xHmiCloseSafetyDoor : BOOL; // Импульс ручного закрытия операторской двери
	xHmiOpenHatch       : BOOL; // Импульс ручного открытия роботного люка
	xHmiCloseHatch      : BOOL; // Импульс ручного закрытия роботного люка
	xHmiUnlockHatch     : BOOL; // Импульс ручного открытия замка роботного люка
	xHmiLockHatch       : BOOL; // Импульс ручного закрытия замка роботного люка
	xHmiOpenChuck       : BOOL; // Импульс ручного разжима патрона
	xHmiCloseChuck      : BOOL; // Импульс ручного зажима патрона
	xHmiSetBlank	  : BOOL; // Ручное подтверждение загруженной заготовки
    xHmiSetDetail     : BOOL; // Ручное подтверждение загруженной детали
	xHmiEnable        : BOOL; // Импульс включения станка или отмены ожидающего отключения
	xHmiDisable       : BOOL; // Импульс отключения станка от работы
	xHmiAcceptRunCNC  : BOOL; // Импульс подтверждения запуска цикла обработки на станке 
	xHmiRejectRunCNC  : BOOL; // Импульс отклонения запуска цикла обработки на станке
	xHmiAcceptDoor    : BOOL; // Импульс подтверждения оператора закрытии двери
	xHmiRejectDoor    : BOOL; // Импульс отклонения оператора закрытии двери
	xUseHmiCycleTime  : BOOL; // TRUE: использовать время цикла, заданное с HMI
	tHmiCycleTime     : TIME; // Начальная или постоянная оценка времени цикла
	stTimeouts        : ST_MACHINE_TIMEOUTS; // Настраиваемые таймауты технологического автомата
	stChangeRecipe    : ARRAY [0..40] OF ST_MACHINE_RECIPE; // Рецепт смены детали
	stLoadRecipe      : ARRAY [0..40] OF ST_MACHINE_RECIPE; // Рецепт загрузки заготовки
	stUnloadRecipe    : ARRAY [0..40] OF ST_MACHINE_RECIPE; // Рецепт выгрузки детали
	stPoints          : ST_MACHINE_POINTS; // Имена рабочих точек станка
	stRobotStatus     : ST_ROBOT_STATUS; // Статусы робота
	eRobotTargetPoint : E_POINT_NAME; // Защёлкнутая текущая цель робота
	stMachineStatus   : ST_MACHINE_IO_STATUS; // Состояние исполнительных механизмов станка
END_VAR
VAR_OUTPUT
	Command : ST_MACHINE_COMMAND; // Команды станку и роботу
	Status  : ST_MACHINE_PUBLIC; // Публичные статусы станка
	Diag    : ST_MACHINE_DIAG; // Состояние автомата и выбранная операция
	Error   : ST_MACHINE_ERRORS; // Активные и последние ошибки
END_VAR
VAR
	eState                  : E_MACHINE_STATE := E_MACHINE_STATE.DISABLED; // Текущее состояние автомата
	ePartState              : E_PART_STATE := E_PART_STATE.UNKNOWN; // Состояние детали в патроне
	ePartType               : E_PART_TYPE := E_PART_TYPE.UNKNOWN; // Тип детали в патроне 
	uiIndex                 : UINT; // Индекс команды рецепта
	tofErrorDoor            : TOF; // Контроль закрытия люка при нахождении робота внутри
	rtExectue               : R_TRIG; // Фронт команды запуска
	rtEnabledMachine        : R_TRIG; // Фронт команды включения
	rtDisabledMachine       : R_TRIG; // Фронт команды отключения
	rtResetMachine          : R_TRIG; // Фронт локального или общего сброса ошибки станка
	rtCycleDone             : R_TRIG; // Фронт завершения цикла станка
	rtCycleStarted          : R_TRIG; // Фронт фактического запуска обработки
	ftCycleStopped          : F_TRIG; // Спад фактического цикла обработки
	rtSetBlankLoaded        : R_TRIG; // Фронт ручного подтверждения заготовки
    rtSetDetailLoaded       : R_TRIG; // Фронт ручного подтверждения детали
	rtHmiOpenSafetyDoor      : R_TRIG; // Фронт ручного открытия операторской двери
	rtHmiCloseSafetyDoor     : R_TRIG; // Фронт ручного закрытия операторской двери
	rtHmiOpenHatch           : R_TRIG; // Фронт ручного открытия люка
	rtHmiCloseHatch          : R_TRIG; // Фронт ручного закрытия люка
	rtHmiUnlockHatch         : R_TRIG; // Фронт ручного открытия замка
	rtHmiLockHatch           : R_TRIG; // Фронт ручного закрытия замка
	rtDoorClosed             : R_TRIG; // Фронт подтверждённого закрытия роботного люка
	rtHmiOpenChuck           : R_TRIG; // Фронт ручного разжима патрона
	rtHmiCloseChuck          : R_TRIG; // Фронт ручного зажима патрона
	ftChuckClamped          : F_TRIG; // Спад закрытия кулачков
	tonCycleMeasure         : TON; // Измерение длительности автоматического цикла
	tonRobotMoveTimeout     : TON; // Ограничение времени перемещения робота
	tonRobotActionTimeout   : TON; // Ограничение времени действия захвата
	tonRobotReleaseTimeout  : TON; // Ограничение времени освобождения интерфейса робота
	tonDoorOpenTimeout      : TON; // Ограничение времени открытия двери
	tonDoorCloseTimeout     : TON; // Ограничение времени закрытия двери
	tonHatchUnlockTimeout   : TON; // Ограничение времени открытия замка
	tonChuckOpenTimeout     : TON; // Ограничение времени разжима патрона
	tonChuckCloseTimeout    : TON; // Ограничение времени зажима патрона
	tonCycleStartTimeout    : TON; // Ограничение времени подтверждения запуска цикла
	xOperatorRunningCNC     : BOOL; // Оператор запустил цикл обработки с панели оператора
	xOperatorClosingDoor    : BOOL; // Оператор запустил закрытие дверей
	xAutoCycleCommanded     : BOOL; // Цикл был запущен этим блоком
	xCycleMeasureActive     : BOOL; // Измеряется текущий автоматический цикл
	xCycleMeasureValid      : BOOL; // Текущее измерение можно сохранить
	xMeasuredTimeValid      : BOOL; // Получено корректное измеренное время
	tMeasuredCycle          : TIME; // Последнее корректное измеренное время
	tExpectedCycle          : TIME; // Ожидаемое время текущего цикла
	xRetreatStarted         : BOOL; // Начат отход робота от станка
	xRobotInsideMachine     : BOOL; // Робот находится внутри рабочей зоны
	xFaultContextCaptured   : BOOL; // Контекст робота зафиксирован при входе в ERROR
	xRobotInsideAtFault     : BOOL; // Робот был в зоне станка при возникновении ошибки
	xDoorRobotStopLatched  : BOOL; // Останов по люку удерживается до полной остановки Motion
	xRobotStopRequired      : BOOL; // Итоговая реакция ROBOT_STOP, сформированная станком
	xRobotResetDependencyReady : BOOL; // Каскадная ошибка робота может быть сброшена тем же импульсом
	xDoorRobotRecoveryReady : BOOL; // Люк открыт либо робот уже вышел из рабочей зоны
	xManualHatchRecoveryOpenAllowed : BOOL; // Разрешено открыть люк для безопасного восстановления
	xSafetyDoorSafe        : BOOL; // Оба сигнала операторской двери непротиворечиво подтверждают закрытие
	xManualControlAllowed  : BOOL; // Общие условия ручного управления механизмами
	xManualSafetyDoorOpenAllowed  : BOOL;
	xManualSafetyDoorCloseAllowed : BOOL;
	xManualHatchOpenAllowed       : BOOL;
	xManualHatchCloseAllowed      : BOOL;
	xManualHatchUnlockAllowed     : BOOL;
	xManualHatchLockAllowed       : BOOL;
	xManualChuckOpenAllowed       : BOOL;
	xManualChuckCloseAllowed      : BOOL;
	xRobotDone              : BOOL; // Робот освобождён алгоритмом станка
	xServiceDoorCloseDemand : BOOL; // Внутренний запрос закрытия двери
	xServiceDoorOpenDemand  : BOOL; // Внутренний запрос открытия двери
	xServiceHatchUnlockDemand : BOOL; // Внутренний запрос открытия замка
	xManualHatchUnlockDemand  : BOOL; // Защёлкнутое ручное состояние открытия замка
	xManualHatchOpenDemand    : BOOL; // Ручное открытие люка после снятия замка
	xAutoDoorOpenLatched    : BOOL; // Защёлка автоматического открытия двери
	xRobotActionDone        : BOOL; // Запрошенное действие захвата уже выполнено
	xRobotCommandStarted    : BOOL; // Текущий шаг рецепта действительно принят FB_ROBOT
	xDisableRequest         : BOOL; // Сохранённый запрос отключения после операции или обработки
	eGrantedOperation       : E_MACHINE_OPERATION; // Разрешённая операция обслуживания
	eActualOperation        : E_MACHINE_OPERATION; // Выполняемая операция обслуживания
	stRecipe                : ARRAY [0..40] OF ST_MACHINE_RECIPE; // Активный рецепт операции
END_VAR

VAR CONSTANT
	ERR_WRONG_OPERATION     : DWORD := 1;       // Выбрана неподдерживаемая операция
	ERR_WRONG_COMMAND       : DWORD := 2;       // В рецепте встретился неподдерживаемый шаг
	ERR_ROBOT_MOTION        : DWORD := 4;       // Робот перешёл в ошибку при движении
	ERR_ROBOT_ACTION        : DWORD := 8;       // Робот перешёл в ошибку при действии захвата
	ERR_DOOR_OPEN           : DWORD := 16;      // Авария станка при открытии люка
	ERR_DOOR_CLOSE          : DWORD := 32;      // Авария станка при закрытии люка
	ERR_CHUCK_OPEN          : DWORD := 64;      // Авария станка при разжиме патрона
	ERR_CHUCK_CLOSE         : DWORD := 128;     // Авария станка при зажиме патрона
	ERR_CYCLE_START         : DWORD := 256;     // Авария станка при запуске цикла
	ERR_SAFETY_STOP         : DWORD := 512;     // Глобальная ошибка ячейки
	ERR_UNKNOWN_DETAIL      : DWORD := 1024;    // Неизвестно содержимое патрона
	ERR_MACHINE_ALARM       : DWORD := 2048;    // Физическая авария станка
	ERR_INDEX               : DWORD := 4096;    // Индекс рецепта вышел за диапазон
	ERR_DOOR_ROBOT          : DWORD := 8192;    // Люк закрывается при роботе в зоне
	ERR_MACHINE_IDLE        : DWORD := 16384;   // Физическая авария станка в IDLE
	ERR_TIMEOUT_ROBOT_MOVE    : DWORD := DWORD#16#00008000; // Таймаут перемещения робота
	ERR_TIMEOUT_ROBOT_ACTION  : DWORD := DWORD#16#00010000; // Таймаут действия захвата
	ERR_TIMEOUT_ROBOT_RELEASE : DWORD := DWORD#16#00020000; // Таймаут освобождения интерфейса робота
	ERR_TIMEOUT_DOOR_OPEN     : DWORD := DWORD#16#00040000; // Таймаут открытия двери
	ERR_TIMEOUT_DOOR_CLOSE    : DWORD := DWORD#16#00080000; // Таймаут закрытия двери
	ERR_TIMEOUT_CHUCK_OPEN    : DWORD := DWORD#16#00100000; // Таймаут разжима патрона
	ERR_TIMEOUT_CHUCK_CLOSE   : DWORD := DWORD#16#00200000; // Таймаут зажима патрона
	ERR_TIMEOUT_CYCLE_START   : DWORD := DWORD#16#00400000; // Таймаут подтверждения запуска цикла
	ERR_SAFETY_DOOR_OPEN     : DWORD := DWORD#16#00800000; // Дверь открылась во время обслуживания
	ERR_TIMEOUT_HATCH_UNLOCK : DWORD := DWORD#16#01000000; // Таймаут открытия замка роботного люка
	ERR_HATCH_UNLOCK_PROCESSING : DWORD := DWORD#16#02000000; // Замок открыт во время обработки

	// Эти ошибки уже относятся к действию робота и всегда имеют эффект ROBOT_STOP.
	MASK_ALWAYS_ROBOT_STOP : DWORD :=
								ERR_ROBOT_MOTION OR
								ERR_ROBOT_ACTION OR
								ERR_DOOR_ROBOT OR
								ERR_SAFETY_DOOR_OPEN OR
								ERR_TIMEOUT_ROBOT_MOVE OR
								ERR_TIMEOUT_ROBOT_ACTION OR
								ERR_TIMEOUT_ROBOT_RELEASE;

	// Первичные ошибки станка: EQUIPMENT_STOP без робота и ROBOT_STOP с роботом.
	MASK_EQUIPMENT_ERROR : DWORD :=
								ERR_WRONG_OPERATION OR
								ERR_WRONG_COMMAND OR
								ERR_DOOR_OPEN OR
								ERR_DOOR_CLOSE OR
								ERR_CHUCK_OPEN OR
								ERR_CHUCK_CLOSE OR
								ERR_CYCLE_START OR
								ERR_UNKNOWN_DETAIL OR
								ERR_MACHINE_ALARM OR
								ERR_INDEX OR
								ERR_MACHINE_IDLE OR
								ERR_TIMEOUT_DOOR_OPEN OR
								ERR_TIMEOUT_DOOR_CLOSE OR
								ERR_TIMEOUT_CHUCK_OPEN OR
								ERR_TIMEOUT_CHUCK_CLOSE OR
								ERR_TIMEOUT_CYCLE_START OR
								ERR_TIMEOUT_HATCH_UNLOCK OR
								ERR_HATCH_UNLOCK_PROCESSING;
								
	// Ошибки, полученные от других блоков или общей логики ячейки.
	MASK_EXTERNAL_ERROR  	: DWORD :=
								ERR_SAFETY_STOP OR
								ERR_ROBOT_ACTION OR
								ERR_ROBOT_MOTION;

	WRN_RESET_ALARM_ACTIVE : UINT := 1; // Сброс отклонён из-за физической аварии станка
	WRN_RESET_GLOBAL_ERROR : UINT := 2; // Сброс отклонён из-за глобальной ошибки
	WRN_RESET_EXECUTE      : UINT := 3; // Сброс отклонён во время операции обслуживания
	WRN_ENABLE_ALARM_ACTIVE: UINT := 4; // Включение отклонено из-за физической аварии станка
	WRN_ENABLE_PROCESSING  : UINT := 5; // Включение отклонено во время обработки
	WRN_ENABLE_PART_UNKNOWN: UINT := 7; // Состояние изделия в патроне не определено
	WRN_RESET_ROBOT_ERROR  : UINT := 8; // Каскадная ошибка робота ещё не готова к сбросу
	WRN_ENABLE_SAFETY_DOOR_OPEN : UINT := 9; // Включение отклонено: операторская дверь не закрыта
	WRN_MANUAL_CONTROL_REJECTED : UINT := 10; // Ручная команда механизма отклонена PLC
	WRN_ENABLE_POINTS : UINT := 11; // Не настроены рабочие точки этого станка
							
	
END_VAR

rtEnabledMachine (CLK :=xHmiEnable);
rtDisabledMachine (CLK :=xHmiDisable);
rtResetMachine(CLK := xReset OR xResetGlobal);
rtCycleDone(CLK := stMachineStatus.xCycleDone);
rtCycleStarted(CLK := stMachineStatus.xCycleActive);
ftCycleStopped(CLK := stMachineStatus.xCycleActive);
rtSetBlankLoaded(CLK := xHmiSetBlank);
rtSetDetailLoaded(CLK := xHmiSetDetail);
rtHmiOpenSafetyDoor(CLK := xHmiOpenSafetyDoor);
rtHmiCloseSafetyDoor(CLK := xHmiCloseSafetyDoor);
rtHmiOpenHatch(CLK := xHmiOpenHatch);
rtHmiCloseHatch(CLK := xHmiCloseHatch);
rtHmiUnlockHatch(CLK := xHmiUnlockHatch);
rtHmiLockHatch(CLK := xHmiLockHatch);
rtDoorClosed(CLK := stMachineStatus.xDoorClosed);
rtHmiOpenChuck(CLK := xHmiOpenChuck);
rtHmiCloseChuck(CLK := xHmiCloseChuck);
ftChuckClamped(CLK := stMachineStatus.xChuckClamped);

xSafetyDoorSafe := stMachineStatus.xSafetyDoorClosed
	AND NOT stMachineStatus.xSafetyDoorOpen;

// Считаем робота находящимся в зоне также по активной цели: текущая точка
// обновляется только после завершения движения и иначе пропускает закрытие
// люка в последнем участке маршрута.
xRobotInsideMachine := (eState = E_MACHINE_STATE.ROBOT_ACTION)
	OR ((eState = E_MACHINE_STATE.ROBOT_MOVE)
		AND (stRecipe[uiIndex].stPoint <> E_MACHINE_POINTS.ABOVE))
	OR (stRobotStatus.eCurrentPoint = stPoints.eInside)
	OR (stRobotStatus.eCurrentPoint = stPoints.eChuck)
	OR (stRobotStatus.eCurrentPoint = stPoints.eChuckApproach)
	OR (stRobotStatus.xBusy
		AND ((eRobotTargetPoint = stPoints.eInside)
			OR (eRobotTargetPoint = stPoints.eChuck)
			OR (eRobotTargetPoint = stPoints.eChuckApproach)))
	// FB_ROBOT очищает eActivePoint сразу после принятого Stop. Пока
	// аварийная защёлка не отпущена, считаем робота оставшимся внутри зоны.
	OR xDoorRobotStopLatched;

// Ручное управление разрешено только при выбранном ручном режиме и остановленном
// автомате станка. xAutomaticUseEnabled хранит выбор для следующей автообработки
// и не является текущим владельцем станка: после аварии и сброса этот флаг
// остаётся TRUE, хотя eState уже DISABLED и автоматикой станок не управляется.
// Конкретные xAllowed дополнительно не дают отправлять бессмысленную команду
// уже достигнутого положения.
xManualControlAllowed := xManualMode
	AND NOT xIoManual
	AND (eState = E_MACHINE_STATE.DISABLED)
	AND NOT xGlobalError
	AND NOT stMachineStatus.xAlarm
	AND NOT stMachineStatus.xCycleActive;

// После аварии «робот внутри/люк закрыт» разрешается только открыть люк,
// причём лишь после полной остановки Motion-слоя. Остальные механизмы остаются
// заблокированы до штатного сброса ошибки.
xDoorRobotRecoveryReady := (stMachineStatus.xDoorOpen AND NOT stMachineStatus.xDoorClosed)
	OR NOT xRobotInsideMachine;
xManualHatchRecoveryOpenAllowed := xManualMode
	AND NOT xIoManual
	AND (eState = E_MACHINE_STATE.ERROR)
	AND ((Error.dwErrorActive AND ERR_DOOR_ROBOT) <> DWORD#0)
	AND stMachineStatus.xDoorClosed
	AND NOT stMachineStatus.xDoorOpen
	AND NOT stMachineStatus.xAlarm
	AND NOT stMachineStatus.xCycleActive
	AND xSafetyDoorSafe
	AND NOT xGlobalError
	AND NOT xRobotMotionBusy
	AND NOT stRobotStatus.xBusy;
xManualSafetyDoorOpenAllowed := xManualControlAllowed AND xSafetyDoorControlEnabled
	AND stMachineStatus.xSafetyDoorClosed
	AND NOT stMachineStatus.xSafetyDoorOpen;
xManualSafetyDoorCloseAllowed := xManualControlAllowed AND xSafetyDoorControlEnabled
	AND stMachineStatus.xSafetyDoorOpen
	AND NOT stMachineStatus.xSafetyDoorClosed;
xManualHatchOpenAllowed := (xManualControlAllowed OR xManualHatchRecoveryOpenAllowed)
	AND stMachineStatus.xDoorClosed
	AND NOT stMachineStatus.xDoorOpen;
xManualHatchCloseAllowed := xManualControlAllowed
	AND stMachineStatus.xDoorOpen
	AND NOT stMachineStatus.xDoorClosed
	AND NOT xRobotInsideMachine;
xManualHatchUnlockAllowed := xManualControlAllowed
	AND stMachineStatus.xDoorClosed
	AND NOT stMachineStatus.xDoorOpen
	AND stMachineStatus.xHatchLocked;
xManualHatchLockAllowed := xManualControlAllowed
	AND NOT stMachineStatus.xHatchLocked
	AND stMachineStatus.xDoorClosed
	AND NOT stMachineStatus.xDoorOpen;
xManualChuckOpenAllowed := xManualControlAllowed
	AND stMachineStatus.xChuckClamped
	AND NOT stMachineStatus.xChuckUnclamped;
xManualChuckCloseAllowed := xManualControlAllowed
	AND stMachineStatus.xChuckUnclamped
	AND NOT stMachineStatus.xChuckClamped;

xRobotResetDependencyReady := (((Error.dwErrorActive
		AND MASK_ALWAYS_ROBOT_STOP) = DWORD#0)
		AND (((Error.dwErrorActive AND MASK_EQUIPMENT_ERROR) = DWORD#0)
			OR NOT xRobotInsideAtFault))
	OR NOT stRobotStatus.xError
	OR stRobotStatus.xResetAllowed;

// Любой сброс формирует одно предупреждение с конкретной причиной отказа.
IF rtResetMachine.Q
AND (eState = E_MACHINE_STATE.ERROR) THEN
	IF stMachineStatus.xAlarm THEN
		Diag.stWarning.uiCode := WRN_RESET_ALARM_ACTIVE;
	ELSIF xGlobalError THEN
		Diag.stWarning.uiCode := WRN_RESET_GLOBAL_ERROR;
	ELSIF xExecute THEN
		Diag.stWarning.uiCode := WRN_RESET_EXECUTE;
	ELSIF ((Error.dwErrorActive AND ERR_DOOR_ROBOT) <> DWORD#0)
	AND NOT xDoorRobotRecoveryReady THEN
		Diag.stWarning.uiCode := WRN_RESET_ROBOT_ERROR;
	ELSIF NOT xRobotResetDependencyReady THEN
		Diag.stWarning.uiCode := WRN_RESET_ROBOT_ERROR;
	ELSE
		Diag.stWarning.uiCode := UINT#0;
	END_IF;

	IF Diag.stWarning.uiCode <> UINT#0 THEN
		Diag.stWarning.udiSequence := Diag.stWarning.udiSequence + UDINT#1;
		IF Diag.stWarning.udiSequence = UDINT#0 THEN
			Diag.stWarning.udiSequence := UDINT#1;
		END_IF;
	END_IF;
END_IF;

// Отклонённая попытка включения регистрируется в журнале предупреждений.
IF rtEnabledMachine.Q
AND (eState = E_MACHINE_STATE.DISABLED)
AND (stMachineStatus.xAlarm
	OR stMachineStatus.xCycleActive
	OR NOT xSafetyDoorSafe
	OR NOT xPointsConfigured
	OR (ePartState = E_PART_STATE.UNKNOWN)) THEN
	IF NOT xPointsConfigured THEN
		Diag.stWarning.uiCode := WRN_ENABLE_POINTS;
	ELSIF stMachineStatus.xAlarm THEN
		Diag.stWarning.uiCode := WRN_ENABLE_ALARM_ACTIVE;
	ELSIF stMachineStatus.xCycleActive THEN
		Diag.stWarning.uiCode := WRN_ENABLE_PROCESSING;
	ELSIF NOT xSafetyDoorSafe THEN
		Diag.stWarning.uiCode := WRN_ENABLE_SAFETY_DOOR_OPEN;
	ELSE
		Diag.stWarning.uiCode := WRN_ENABLE_PART_UNKNOWN;
	END_IF;

	Diag.stWarning.udiSequence := Diag.stWarning.udiSequence + UDINT#1;
	IF Diag.stWarning.udiSequence = UDINT#0 THEN
		Diag.stWarning.udiSequence := UDINT#1;
	END_IF;
END_IF;

// HMI показывает xAllowed только визуально. Любая фактически отклонённая
// команда всё равно фиксируется PLC-предупреждением и попадает в журнал.
IF (rtHmiOpenSafetyDoor.Q AND NOT xManualSafetyDoorOpenAllowed)
OR (rtHmiCloseSafetyDoor.Q AND NOT xManualSafetyDoorCloseAllowed)
OR (rtHmiOpenHatch.Q AND NOT xManualHatchOpenAllowed)
OR (rtHmiCloseHatch.Q AND NOT xManualHatchCloseAllowed)
OR (rtHmiUnlockHatch.Q AND NOT xManualHatchUnlockAllowed)
OR (rtHmiLockHatch.Q AND NOT xManualHatchLockAllowed)
OR (rtHmiOpenChuck.Q AND NOT xManualChuckOpenAllowed)
OR (rtHmiCloseChuck.Q AND NOT xManualChuckCloseAllowed) THEN
	Diag.stWarning.uiCode := WRN_MANUAL_CONTROL_REJECTED;
	Diag.stWarning.udiSequence := Diag.stWarning.udiSequence + UDINT#1;
	IF Diag.stWarning.udiSequence = UDINT#0 THEN
		Diag.stWarning.udiSequence := UDINT#1;
	END_IF;
END_IF;

// Повторное включение отменяет ещё не выполненный запрос отключения.
// Одновременным командам отдаётся безопасный приоритет отключения.
IF rtDisabledMachine.Q THEN
	xDisableRequest := TRUE;
ELSIF rtEnabledMachine.Q AND xDisableRequest THEN
	xDisableRequest := FALSE;
END_IF;

// Измеряются только циклы, запущенные автоматикой этого блока.
IF rtCycleStarted.Q THEN
	xCycleMeasureActive := xAutoCycleCommanded;
	xCycleMeasureValid := xAutoCycleCommanded;
END_IF;

IF xCycleMeasureActive
AND (stMachineStatus.xAlarm
	OR xGlobalError
	OR (eState = E_MACHINE_STATE.ERROR)
	OR (eState = E_MACHINE_STATE.DISABLED)) THEN
	xCycleMeasureValid := FALSE;
END_IF;

IF ftCycleStopped.Q THEN
	IF xCycleMeasureActive
	AND xCycleMeasureValid
	AND (tonCycleMeasure.ET > T#0S) THEN
		tMeasuredCycle := tonCycleMeasure.ET;
		xMeasuredTimeValid := TRUE;
	END_IF;
	xCycleMeasureActive := FALSE;
	xCycleMeasureValid := FALSE;
	xAutoCycleCommanded := FALSE;
END_IF;

tonCycleMeasure(
	IN := stMachineStatus.xCycleActive,
	PT := T#24H
);

// Таймеры работают только в исполнительных шагах. При переходе в другой шаг
// соответствующий экземпляр TON сбрасывается автоматически.
tonRobotMoveTimeout(
	IN := eState = E_MACHINE_STATE.ROBOT_MOVE,
	PT := stTimeouts.tRobotMove
);
tonRobotActionTimeout(
	IN := eState = E_MACHINE_STATE.ROBOT_ACTION,
	PT := stTimeouts.tRobotAction
);
tonRobotReleaseTimeout(
	IN := eState = E_MACHINE_STATE.RELEASE_ROBOT_ACTION,
	PT := stTimeouts.tRobotRelease
);
tonDoorOpenTimeout(
	IN := eState = E_MACHINE_STATE.DOOR_OPEN,
	PT := stTimeouts.tDoorOpen
);
tonDoorCloseTimeout(
	IN := eState = E_MACHINE_STATE.DOOR_CLOSE,
	PT := stTimeouts.tDoorClose
);
tonHatchUnlockTimeout(
	IN := (eState <> E_MACHINE_STATE.ERROR)
		AND stMachineStatus.xHatchLocked
		AND (((eState = E_MACHINE_STATE.DOOR_OPEN) AND xServiceHatchUnlockDemand)
			OR (xManualHatchUnlockDemand AND xManualMode)),
	PT := stTimeouts.tHatchUnlock
);
tonChuckOpenTimeout(
	IN := eState = E_MACHINE_STATE.CHUCK_OPEN,
	PT := stTimeouts.tChuckOpen
);
tonChuckCloseTimeout(
	IN := eState = E_MACHINE_STATE.CHUCK_CLOSE,
	PT := stTimeouts.tChuckClose
);
tonCycleStartTimeout(
	IN := eState = E_MACHINE_STATE.CYCLE_START,
	PT := stTimeouts.tCycleStart
);

// В автоматическом режиме до первого измерения используется время с HMI.
IF xUseHmiCycleTime THEN
	tExpectedCycle := tHmiCycleTime;
ELSIF xMeasuredTimeValid THEN
	tExpectedCycle := tMeasuredCycle;
ELSE
	tExpectedCycle := tHmiCycleTime;
END_IF;

